(* IEC 61131-3 sources: plcassist-cli/packages/volt-lsp-iec/test-corpus/lenze-mid/Device/Plc Logic/Application/Library Manager/L_CT1P_ControlToolbox, 48 files *)

(* ---- L_CT1P_CONSTANTS.gvl ---- *)
VAR_GLOBAL
	GCWFRICTIONHISTMAX : WORD := 99;
	GCMAXPARITEMS : WORD := 35;
	GCPARITEMSUSED : WORD := 34;
END_VAR

(* ---- L_CT1P_INTERNALCONST.gvl ---- *)
VAR_GLOBAL
END_VAR

(* ---- L_CT1P_IKINAUTOTUNINGEXTERNAL.itf ---- *)
INTERFACE L_CT1P_IKINAUTOTUNINGEXTERNAL
END_INTERFACE

METHOD CALLDEVICEPARAMMANAGERSLAVE
VAR_INPUT
	ECOMMAND : WORD;
	WREGISTERPOSITION : WORD;
	XEXECUTE : BOOL;
END_VAR
VAR_OUTPUT
	XBUSY : BOOL;
	XDONE : BOOL;
	XERROR : BOOL;
	EERRORID : L_Ie1P_Error;
END_VAR
END_METHOD

METHOD CALLMONITORING : BOOL
VAR_INPUT
	XENABLE : BOOL;
END_VAR
END_METHOD

METHOD CHECKPRECONDITIONS : WORD
VAR_INPUT
	XENABLE : BOOL;
	PSCAUTOTUNINGDATAMAININ : POINTER TO BYTE;
END_VAR
END_METHOD

METHOD CLOSEBRAKESPEEDINDEPENDET
VAR_INPUT
	XCLOSBRAKESPEEDINDEPENDET : BOOL;
END_VAR
END_METHOD

METHOD GETMAINFOLLOWERAXIS
VAR_OUTPUT
	PMAINAXISOUT : POINTER TO AXIS_REF;
	PFOLLOWINGAXISOUT : POINTER TO AXIS_REF;
END_VAR
END_METHOD

METHOD SPEEDEQUALSZERO : BOOL
END_METHOD

METHOD STORESAMPLEDBRAKETORQUE
VAR_INPUT
	XSTOREVALUE : BOOL;
END_VAR
END_METHOD

(* ---- _TXERROR.fun ---- *)
FUNCTION _TXERROR : L_IE1P_Error
VAR_INPUT
	WERRCODE : WORD;
END_VAR
END_FUNCTION

(* ---- GETBOOLEANPROPERTY.fun ---- *)
FUNCTION GETBOOLEANPROPERTY : BOOL
VAR_INPUT
	STKEY : WSTRING;
END_VAR
END_FUNCTION

(* ---- GETCOMPANY.fun ---- *)
FUNCTION GETCOMPANY : WSTRING
END_FUNCTION

(* ---- GETNUMBERPROPERTY.fun ---- *)
FUNCTION GETNUMBERPROPERTY : DINT
VAR_INPUT
	STKEY : WSTRING;
END_VAR
END_FUNCTION

(* ---- GETTEXTPROPERTY.fun ---- *)
FUNCTION GETTEXTPROPERTY : WSTRING
VAR_INPUT
	STKEY : WSTRING;
END_VAR
END_FUNCTION

(* ---- GETTEXTPROPERTY2.fun ---- *)
FUNCTION GETTEXTPROPERTY2 : POINTER TO WSTRING
VAR_INPUT
	STKEY : WSTRING;
END_VAR
END_FUNCTION

(* ---- GETTITLE.fun ---- *)
FUNCTION GETTITLE : WSTRING
END_FUNCTION

(* ---- GETVERSION.fun ---- *)
FUNCTION GETVERSION : VERSION
END_FUNCTION

(* ---- GETVERSIONPROPERTY.fun ---- *)
FUNCTION GETVERSIONPROPERTY : VERSION
VAR_INPUT
	STKEY : WSTRING;
END_VAR
END_FUNCTION

(* ---- L_CT1P_CA_CALCDISTANCE.fun ---- *)
FUNCTION L_CT1P_CA_CALCDISTANCE : BOOL
VAR_INPUT
	LRCONSTVELTIME : LREAL;
	LRVELOCITYMAX : LREAL;
	LRACCDECMAX : LREAL;
END_VAR
VAR_OUTPUT
	XERROR : BOOL;
	EERRORID : L_IE1P_Error;
	LRTARGETPOSRELATIVEINT : LREAL;
END_VAR
END_FUNCTION

(* ---- L_CT1P_CA_CALCPROFILEPARAMS.fun ---- *)
FUNCTION L_CT1P_CA_CALCPROFILEPARAMS : BOOL
VAR_INPUT
	LRMAXVELOCITYIN : LREAL := 0;
	LRMAXACCELERATIONIN : LREAL := 0;
	LRMAXDISTANCEIN : LREAL := 0;
END_VAR
VAR_OUTPUT
	LRVELOCITYACTIVE : LREAL := 0;
	LRACCELERATIONACTIVE : LREAL := 0;
	LRMOVEMENTDISTANCEMIN : LREAL := 0;
	LRMOVEMENTDISTANCEMAX : LREAL := 0;
	LRCONSTVELTIME : LREAL := 0;
END_VAR
END_FUNCTION

(* ---- L_CT1P_CA_GETTIMINGOFEXTERNALENCODER.fun ---- *)
FUNCTION L_CT1P_CA_GETTIMINGOFEXTERNALENCODER : BOOL
VAR_OUTPUT
	LRDELAYACTPOS : LREAL;
	LRFILTERCYCLESACTPOS : LREAL;
END_VAR
VAR_IN_OUT
	REALAXIS : _Axis_Ref_Real;
END_VAR
END_FUNCTION

(* ---- L_CT1P_CHECKBASEVALUES.fun ---- *)
FUNCTION L_CT1P_CHECKBASEVALUES : WORD
VAR_INPUT
	PSCCOREDATA : POINTER TO L_CT1P_CA_DeviceParamList;
END_VAR
VAR_IN_OUT
	AXIS : AXIS_REF;
END_VAR
END_FUNCTION

(* ---- L_CT1P_GETOCCOMPDELTAPOSITION.fun ---- *)
FUNCTION L_CT1P_GETOCCOMPDELTAPOSITION : LREAL
VAR_INPUT
	LREIGENFREQ : LREAL;
	LRAMPRATIO : LREAL;
	ECOMPMODE : L_CT1P_OscCompMode;
	LRTARGETVELOCITY : LREAL;
END_VAR
END_FUNCTION

(* ---- L_CT1P_GETOCCOMPDELTATIME.fun ---- *)
FUNCTION L_CT1P_GETOCCOMPDELTATIME : LREAL
VAR_INPUT
	LREIGENFREQ : LREAL;
	ECOMPMODE : L_CT1P_OscCompMode;
END_VAR
END_FUNCTION

(* ---- GLOBALTEXTLIST.fb ---- *)
FUNCTION_BLOCK GLOBALTEXTLIST
VAR
	M_TEXTLISTFILE : STRING(255);
	_STNAMESPACE : STRING;
END_VAR
END_FUNCTION_BLOCK

(* ---- IMAGEPOOL.fb ---- *)
FUNCTION_BLOCK IMAGEPOOL
VAR
	M_STNAMESPACE : STRING(80);
	M_STHELPVARID : STRING;
	M_STHELPVARPATH : STRING(255);
	M_STHELP : STRING;
	M_REGISTERIMAGES : BOOL := TRUE;
END_VAR
END_FUNCTION_BLOCK

METHOD FB_INIT : BOOL
VAR_INPUT
	BINITRETAINS : BOOL;
	BINCOPYCODE : BOOL;
END_VAR
END_METHOD

METHOD FB_REINIT : BOOL
END_METHOD

METHOD FB_EXIT : BOOL
VAR_INPUT
	BINCOPYCODE : BOOL;
END_VAR
END_METHOD

(* ---- L_CT1P_AT_TON.fb ---- *)
FUNCTION_BLOCK L_CT1P_AT_TON
VAR_INPUT
	IN : BOOL;
	PT : TIME;
	LRCYCLE : LREAL;
END_VAR
VAR_OUTPUT
	Q : BOOL;
	ET : TIME;
END_VAR
VAR
	TON_INT : TON;
	TCYLCE : TIME;
	XNOTFIRSTCYCLE : BOOL := FALSE;
END_VAR
END_FUNCTION_BLOCK

(* ---- L_CT1P_AUTOTUNING.fb ---- *)
FUNCTION_BLOCK L_CT1P_AUTOTUNING EXTENDS L_MC1P_Template
VAR_INPUT
	XENABLE : BOOL := FALSE;
	XABORT : BOOL := FALSE;
	XRESETERROR : BOOL := FALSE;
	XEXECUTEIDENT : BOOL := FALSE;
	XENABLEPOSITIONWINDOW : BOOL := FALSE;
	LRPOSITIONWINDOWNEG : LREAL := 1.0;
	LRPOSITIONWINDOWPOS : LREAL := 1.0;
	LRVELOCITYLIMIT : LREAL := 0.0;
	LRACCELERATIONLIMIT : LREAL := 0.0;
	LRDISTANCE : LREAL := 0;
	XRESTOREPARAM : BOOL := FALSE;
	XUSEAXISPARAMETER : BOOL := FALSE;
	EALLOWEDDIRECTION : L_MC1P_ServiceDirection := L_MC1P_ServiceDirection.both;
END_VAR
VAR_OUTPUT
	XERROR : BOOL := FALSE;
	XWARNING : BOOL := FALSE;
	EERRORID : L_IE1P_Error := L_IE1P_Error.NoError;
	XABORTED : BOOL := FALSE;
	XIDENTBUSY : BOOL := FALSE;
	XIDENTDONE : BOOL := FALSE;
	EIDENTIFICATIONSTATE : L_CT1P_CA_IdentificationState := L_CT1P_CA_IdentificationState.PLC_Reset;
	XPOSITIONWINDOWENABLED : BOOL := FALSE;
	LRMVMTVELMAX : LREAL := 0.0;
	LRMVMTACCMAX : LREAL := 0.0;
	LRMVMTDISTANCEMIN : LREAL := 0;
	LRVPNACT : LREAL := 0.0;
	LRTNNACT : LREAL := 0.0;
	LRVPPACT : LREAL := 0.0;
END_VAR
VAR
	RTRESTOREPARAM : R_TRIG;
	EACTSTATE : DWORD := 0;
	XLEAVESERVICESTATE : BOOL := FALSE;
	XDISABLESEEN : BOOL := FALSE;
	XABORTSEEN : BOOL := FALSE;
	XRESETERROROLD : BOOL;
	WCNT : WORD := 0;
	SCCOREDATA : L_CT1P_CA_CoreData := STRUCT(pFB_Par := ADR(fb_InternalParamFB), pFB_AxisReadError := ADR(fb_ReadError), pFB_AxisPower := ADR(fb_Power), pFB_Autotuning := THIS);
	TONAUTOTUNINGDURATION : L_CT1P_AT_TON := STRUCT(PT := TIME#1440m0s0ms);
	XEVENTEXTERNALPARAMFBACTIVATED : BOOL := FALSE;
	LRVELOCITYLIMITINT : LREAL := 0;
	LRACCELERATIONLIMITINT : LREAL := 0;
	LRDISTANCEINT : LREAL := 0;
	XEXECUTEIDENTOLD : BOOL := FALSE;
	DEVICEPARAMMANAGER : L_CT1P_CA_DeviceParamManager;
	PROFILEGENERATOR : L_CT1P_CA_ProfileGenerator;
	MONITORING : L_CT1P_CA_Monitoring;
	QUALITYCRITERIA : L_CT1P_CA_QualityCriteria;
	CHECKPRECONDITIONS : L_CT1P_CA_CheckPreconditions;
	PERFORMAUTOTUNING : L_CT1P_CA_PerformAutotuning;
	FB_READERROR : MC_ReadAxisError;
	FB_POWER : mc_power;
	FB_INTERNALPARAMFB : L_CT1P_ParAutoTuninginternal;
	PAXISREAL : POINTER TO _Axis_Ref_Real;
	PBRAKE : POINTER TO L_MC1P_BrakeControlBase;
	PREALAXIS : POINTER TO _AXIS_REF_COM := 0;
	XWARNINGOLD : BOOL := FALSE;
	LRIMPROVEMENTFACTOR : LREAL := 0;
	XDEACTIVATEERRORINAXIS : BOOL := FALSE;
	EALLOWEDDIRECTIONINT : L_MC1P_ServiceDirection := L_MC1P_ServiceDirection.both;
	TON_MAGNETISATION : L_CT1P_AT_TON;
	XAUTOTUNINGWASACTIVE : BOOL;
	XNEWSTEPENTRY : BOOL;
	ENEWSTATE : DWORD;
	XABORTEDOLD : BOOL;
	ITFKINAUTOTUNING : L_CT1P_IKinAutoTuningExternal;
	STATUSOLD : BOOL;
	XSERVICESTATESETBYAXISCMD : BOOL;
	SERVICESTATESETBYAXISCMND : BOOL;
END_VAR
END_FUNCTION_BLOCK

METHOD ATGETACCELERATION : LREAL
VAR_INPUT
	LRVELOCITY : LREAL := 0;
	LRACCELERATION : LREAL := 0;
END_VAR
VAR_IN_OUT
	AXIS : AXIS_REF;
END_VAR
END_METHOD

METHOD ATGETVELOCITY : LREAL
VAR_INPUT
	LRVELOCITY : LREAL := 0;
	LRVELOTIYRATIOPCT : LREAL := 0;
END_VAR
VAR_IN_OUT
	AXIS : AXIS_REF;
END_VAR
END_METHOD

METHOD CALCULATEIMPROVEMENTFACTOR : LREAL
END_METHOD

METHOD CALLINNERFBINSTANCES
END_METHOD

METHOD CALLMOTIONBLOCKS
END_METHOD

METHOD COPYINPUTS
VAR_IN_OUT
	AXIS : Axis_Ref;
END_VAR
END_METHOD

METHOD SETEXTERNALAUTOTUNINGITF
VAR_INPUT
	PIKINAUTOTUNINGIN : POINTER TO L_CT1P_IKinAutoTuningExternal;
END_VAR
END_METHOD

METHOD STATEMACHINE
END_METHOD

METHOD _GETLIBVERSIONASSTRING : STRING
END_METHOD

METHOD _SETEXTERNALPARAMFB
VAR_INPUT
	PPARAMFB : POINTER TO L_CT1P_ParAutoTuninginternal;
END_VAR
END_METHOD

METHOD STATE_CHECKPRECONDITIONSFOLLOWINGAXIS : DWORD
VAR_INPUT
	XSTOP : BOOL;
	EACTSTATE : DWORD;
	ENEXTSTATE : DWORD;
	EABORTSTATE : DWORD;
	EERRORSTATE : DWORD;
END_VAR
END_METHOD

METHOD STATE_CHECKPRECONDITIONS : DWORD
VAR_INPUT
	XSTOP : BOOL;
	EACTSTATE : DWORD;
	ENEXTSTATE : DWORD;
	EABORTSTATE : DWORD;
	EERRORSTATE : DWORD;
END_VAR
END_METHOD

METHOD STATE_DOAUTOTUNE : DWORD
VAR_INPUT
	XSTOP : BOOL;
	EACTSTATE : DWORD;
	ENEXTSTATE : DWORD;
	EABORTSTATE : DWORD;
	EERRORSTATE : DWORD;
END_VAR
END_METHOD

METHOD STATE_FINISH : DWORD
VAR_INPUT
	XSTOP : BOOL;
	EACTSTATE : DWORD;
	ENEXTSTATE : DWORD;
	EABORTSTATE : DWORD;
	EERRORSTATE : DWORD;
END_VAR
END_METHOD

METHOD STATE_PARAMETERHANDLING : DWORD
VAR_INPUT
	XSTOP : BOOL;
	EACTSTATE : DWORD;
	ENEXTSTATE : DWORD;
	EABORTSTATE : DWORD;
	EERRORSTATE : DWORD;
END_VAR
END_METHOD

(* ---- L_CT1P_AXISCOMMAND_AUTOTUNING.fb ---- *)
FUNCTION_BLOCK L_CT1P_AXISCOMMAND_AUTOTUNING EXTENDS L_MC1P_AxisCommand
VAR_INPUT
	PAXIS : POINTER TO AXIS_REF;
END_VAR
VAR
	FB_AUTOTUNING : L_CT1P_Autotuning;
	SCPARAUTOTUNING : REFERENCE TO L_MC1P_AutotuningPara;
	LRCONSTVELTIME : LREAL := 0;
	LRVELOCITYACTIVE : LREAL := 0;
	LRACCELERATIONACTIVE : LREAL := 0;
	LRDISTANCEACTIVE : LREAL := 0;
	SCPARAUTOTUNING_DUMMY : L_MC1P_AutotuningPara;
	PCONNECTOR : POINTER TO IoConfigConnector;
	ITFAXISCOMMMANDAUTOTUNING : L_MC1P_IAxisCommmand_Autotuning;
	AT_FINISHSTATETEMP : WORD := 0;
	EERRORIDTMP : L_IE1P_error := L_IE1P_Error.NoError;
	WMODULETYPE : UINT;
	XDISABLESET : BOOL := FALSE;
	DWINSTANCE : UDINT;
	WNBOFTUNINGDONE : WORD := 1;
	WNBOFEXPECTEDTUNINGS : WORD := 1;
	LRIMPROVEMENTFACTORSTORED : LREAL;
	PBATEXTERNALITF : POINTER TO BYTE;
	PACTIVEAUTOTUNINGAXIS : ARRAY [1..2] OF POINTER TO _AXIS_REF_REAL;
	C_CMDWORKING10 : USINT := 10;
	C_CMDWORKING30 : USINT := 30;
	C_CMDWORKING50 : USINT := 50;
	C_CMDWORKING70 : USINT := 70;
	C_CMDINVALIDTASKCYCLETIME : USINT := 101;
	C_CMDFUNCTIONNOTSUPPORTEDBYFWVERSION : USINT := 104;
	C_CMDPDOINTERFACEDISABLED : USINT := 106;
	C_CMDTESTMODEALREADYACTIVE : USINT := 107;
	C_CMDINVALIDMOTORCONTROLMODE : USINT := 108;
	C_CMDNOVALIDDIRECTION : USINT := 109;
	C_CMDINSTABILITYWITHCHOSENSTRATEGY : USINT := 110;
	C_CMDAXISNOTHOMED : USINT := 111;
	C_AT_STATE_NOTSTARTED : WORD := 0;
	C_AT_STATE_INITIALIZATION : WORD := 1;
	C_AT_STATE_BACKUPDEVICEPARAM : WORD := 2;
	C_AT_STATE_CHECKPRECONDITIONS : WORD := 3;
	C_AT_STATE_AUTOTUNEVPN : WORD := 4;
	C_AT_STATE_AUTOTUNETNN : WORD := 5;
	C_AT_STATE_AUTOTUNEVPP : WORD := 6;
	C_AT_STATE_FINISHED_1 : WORD := 10;
	C_AT_STATE_FINISHED_2 : WORD := 11;
	C_AT_STATE_FINISHED_3 : WORD := 12;
	C_AT_STATE_BACKUPDEVICEPARAMFOLLOWER : WORD := 22;
	C_AT_STATE_CHECKPRECONDITIONSFOLLOWER : WORD := 23;
	C_AT_STATE_AUTOTUNEVPNFOLLOWER : WORD := 24;
	C_AT_STATE_AUTOTUNETNNFOLLOWER : WORD := 25;
	C_AT_STATE_AUTOTUNEVPPFOLLOWER : WORD := 26;
	C_AT_STATE_FINISHED_4 : WORD := 30;
	C_AT_STATE_FINISHED_5 : WORD := 31;
	C_AT_STATE_FINISHED_6 : WORD := 32;
	C_AT_STATE_FINISHED_7 : WORD := 33;
	C_AT_STATE_FINISHED_8 : WORD := 34;
	C_AT_STATE_FINISHED_9 : WORD := 35;
	C_AT_STATE_ABORTING : WORD := 7;
	C_AT_STATE_ABORTEDBYERROR : WORD := 8;
	C_AT_STATE_ABORTEDBYUSER : WORD := 9;
END_VAR
END_FUNCTION_BLOCK

METHOD ABORTING
END_METHOD

METHOD CALCPROFILEPARAMS
VAR_IN_OUT
	AXIS : AXIS_REF;
END_VAR
END_METHOD

METHOD CALCSTATUS
VAR_IN_OUT
	AXIS : _AXIS_REF_REAL;
END_VAR
END_METHOD

METHOD EXECUTE
END_METHOD

METHOD INITIALIZE : UDINT
VAR_INPUT
	WMODULETYPE : UINT;
	DWINSTANCE : UDINT;
	PCONNECTOR : POINTER TO IoConfigConnector;
END_VAR
END_METHOD

METHOD READINPUTS
END_METHOD

METHOD RESETSTATUSPARAMETER
END_METHOD

METHOD UPDATEAXISPOINTER
VAR_INPUT
	PAXIS : POINTER TO AXIS_REF;
END_VAR
END_METHOD

METHOD UPDATEPARAINTERFACE
VAR_IN_OUT
	SCPAR : L_MC1P_AutotuningPara;
END_VAR
END_METHOD

METHOD FB_INIT : BOOL
VAR_INPUT
	BINITRETAINS : BOOL;
	BINCOPYCODE : BOOL;
END_VAR
END_METHOD

(* ---- L_CT1P_BACKLASHCOMP.fb ---- *)
FUNCTION_BLOCK L_CT1P_BACKLASHCOMP EXTENDS L_MC1P_CompensationBase
VAR_INPUT
	LRBACKLASHWIDTH : LREAL := 0.0;
	LRCOMPTIME : LREAL := 0.1;
	ECOMPMODE : L_CT1P_BacklashCompMode := L_CT1P_BacklashCompMode.NegativeComp;
END_VAR
VAR_OUTPUT
	ECONTACTSTATE : L_CT1P_BacklashContactState := L_CT1P_BacklashContactState.Unknown;
END_VAR
VAR
	FBRAMPGEN : L_MC1P_RampGenerator;
	LRBACKLASHWIDTHINT : LREAL;
	LRCOMPTIMEINT : LREAL;
	ECOMPMODEINT : L_CT1P_BacklashCompMode;
	ECOMPREFERENCEINT : L_CT1P_BacklashCompReference;
	LRACCRATIOINT : LREAL := 0.3333333333;
	ECONTACTSTATEINT : L_CT1P_BacklashContactState;
	LRBACKLASHTARGET : LREAL;
	LRBACKLASHTARGETOLD : LREAL;
	LRBACKLASHPOSACT : LREAL;
	LRBACKLASHVELACT : LREAL;
	LRBACKLASHACCACT : LREAL;
	LRBACKLASHPOSOLD : LREAL;
	LRBACKLASHVELOLD : LREAL;
	LRHOMINGOFFSETACT : LREAL;
	LRENABLEPOS : LREAL;
	LRENABLEDIST : LREAL;
	LRENABLEDISTOLD : LREAL;
	LRVELMAX : LREAL;
	LRACCMAX : LREAL;
	ECOMPREFERENCE : L_CT1P_BacklashCompReference := L_CT1P_BacklashCompReference.SetVelocity;
	_CUSTOMINPUTDATA : ARRAY [1..2] OF L_CT1P_BacklashCompInput;
	_CUSTOMOUTPUTDATA : ARRAY [1..2] OF L_CT1P_BacklashCompOutput;
	_PCUSTOMINPUTDATA : POINTER TO L_CT1P_BacklashCompInput;
	_PCUSTOMOUTPUTDATA : POINTER TO L_CT1P_BacklashCompOutput;
	LRACCRATIO : LREAL;
END_VAR
END_FUNCTION_BLOCK

METHOD CALLCYCLIC2
VAR_IN_OUT
	AXIS : Axis_REf;
END_VAR
END_METHOD

METHOD READINPUTS2
VAR_IN_OUT
	AXIS : Axis_REF;
END_VAR
END_METHOD

METHOD RESETOUTPUTS2
VAR_IN_OUT
	AXIS : Axis_REf;
END_VAR
END_METHOD

METHOD CALCULATE2
VAR_IN_OUT
	AXIS : AXIS_REF;
END_VAR
END_METHOD

METHOD CHECKINPUTDATA2
VAR_IN_OUT
	AXIS : Axis_Ref;
END_VAR
END_METHOD

METHOD ENABLEINIT2
VAR_IN_OUT
	AXIS : Axis_REf;
END_VAR
END_METHOD

METHOD LOADOFFSET2
VAR_INPUT
	OFFSET : LREAL;
END_VAR
VAR_IN_OUT
	AXIS : Axis_REf;
END_VAR
END_METHOD

METHOD GETOFFSETVALUES
VAR_OUTPUT
	LROFFSETPOS : LREAL;
	LROFFSETVEL : LREAL;
	LROFFSETACC : LREAL;
END_VAR
END_METHOD

METHOD CALLFUNCTION
VAR_INPUT
	UIINPUTDATAIDX : UINT;
	UIOUTPUTDATAIDX : UINT;
END_VAR
END_METHOD

METHOD COPYINPUTS : BOOL
VAR_INPUT
	IDX : WORD;
END_VAR
END_METHOD

METHOD COPYOUTPUTS : BOOL
VAR_INPUT
	IDX : WORD;
END_VAR
END_METHOD

METHOD GETCOMPTARGET : LREAL
VAR_INPUT
	LRACTBACKLASHTARGET : LREAL;
END_VAR
VAR_IN_OUT
	AXIS : AXIS_REF;
END_VAR
END_METHOD

METHOD GETCONTACTSTATE : L_CT1P_BacklashContactState
VAR_INPUT
	LRBACKLASHWIDTH : LREAL;
	LRBACKLASHPOSACT : LREAL;
	EACTCONTACTSTATE : L_CT1P_BacklashContactState;
END_VAR
VAR_IN_OUT
	AXIS : AXIS_REF;
END_VAR
END_METHOD

METHOD GETDISTANCESINCEENABLE : LREAL
VAR_IN_OUT
	AXIS : AXIS_REF;
END_VAR
END_METHOD

METHOD GETRAMPPARS : BOOL
VAR_INPUT
	LRCOMPTIME : LREAL;
	LRACCRATIO : LREAL;
	LRBACKLASHWIDTH : LREAL;
END_VAR
VAR_OUTPUT
	LRVELMAX : LREAL;
	LRACCMAX : LREAL;
END_VAR
END_METHOD

METHOD GETTRANSDIR : INT
VAR_IN_OUT
	AXIS : AXIS_REF;
END_VAR
END_METHOD

METHOD INITIALIZEFILTER : BOOL
END_METHOD

(* ---- L_CT1P_CA_CHECKPRECONDITIONS.fb ---- *)
FUNCTION_BLOCK L_CT1P_CA_CHECKPRECONDITIONS
VAR_INPUT
	XEXECUTE : BOOL := FALSE;
	XSTOP : BOOL := FALSE;
	RSCCOREDATA : REFERENCE TO L_CT1P_CA_CoreData;
	RDEVICEPARAMMANAGER : REFERENCE TO L_CT1P_CA_DeviceParamManager;
END_VAR
VAR_OUTPUT
	XBUSY : BOOL := FALSE;
	XDONE : BOOL := FALSE;
	XERROR : BOOL := FALSE;
	EERRORID : L_IE1P_Error := L_IE1P_Error.NoError;
END_VAR
VAR_IN_OUT
	AXIS : AXIS_REF;
END_VAR
VAR
	LRSPEEDFILTERTIME : LREAL;
	LRMOTORINERTIA : LREAL;
	LRLOADINERTIA : LREAL;
	RSCACTPARAM : REFERENCE TO L_CT1P_CA_DeviceParam;
	LRVPPREFERENCEVALUE : LREAL;
	LRDELAYACTPOS : LREAL;
	LRFILTERCYCLESACTPOS : LREAL;
	PREALAXIS : POINTER TO _Axis_Ref_Real;
	REALAXIS : REFERENCE TO _Axis_Ref_Real;
	PBRAKE : POINTER TO L_MC1P_BrakeControlBase;
	XSTOPSEEN : BOOL := FALSE;
	XENABLEPROFILECHECK : BOOL;
	DWSTEP : DWORD := 0;
	RTEXECUTE : R_TRIG;
	PROFILECHECK : L_CT1P_CA_ProfileCheck;
END_VAR
END_FUNCTION_BLOCK

METHOD CALLPROFILECHECK
END_METHOD

METHOD CHECKSTOPELSEPROCEEDWITHSTEP
VAR_INPUT
	DWSTEPINP : DWORD;
END_VAR
END_METHOD

METHOD CHECKVALUES : WORD
VAR_IN_OUT
	AXIS : AXIS_REF;
END_VAR
END_METHOD

METHOD RAISEERROR
VAR_INPUT
	ERRCODE : L_IE1P_Error;
END_VAR
END_METHOD

METHOD RAISEFINISHED
END_METHOD

METHOD RAISESTOP
END_METHOD

METHOD READWRITEVALUES : WORD
VAR_IN_OUT
	DWSTEP : DWORD;
	AXIS : AXIS_REF;
END_VAR
END_METHOD

METHOD RESET : BOOL
END_METHOD

METHOD STATEMACHINE
END_METHOD

(* ---- L_CT1P_CA_DEVICEPARAMMANAGER.fb ---- *)
FUNCTION_BLOCK L_CT1P_CA_DEVICEPARAMMANAGER
VAR_INPUT
	ECOMMAND : L_CT1P_CA_DPMCommand := L_CT1P_CA_DPMCommand.None;
	RSCPARAMLIST : REFERENCE TO L_CT1P_CA_DeviceParamList;
	WREGISTERPOSITION : WORD;
	XEXECUTE : BOOL := FALSE;
END_VAR
VAR_OUTPUT
	XBUSY : BOOL := FALSE;
	XDONE : BOOL := FALSE;
	XERROR : BOOL := FALSE;
	EERRORID : L_Ie1P_Error;
END_VAR
VAR_IN_OUT
	AXIS : Axis_ref;
END_VAR
VAR
	WRITEPARAMETER : MC_WriteParameter;
	READPARAMETER : MC_ReadParameter;
	PDCOREAD : POINTER TO L_MC1P.L_DCO_ReadDriveParameter;
	PDCOWRITE : POINTER TO L_MC1P.L_DCO_WriteDriveParameter;
	WWRITEMODE : WORD;
	ECOMMANDINT : L_CT1P_CA_DPMCommand := L_CT1P_CA_DPMCommand.None;
	WREGISTERPOSITIONINT : WORD;
	WIDX : WORD := 1;
	WIDX2 : WORD := 1;
	XEXECUTEOLD : BOOL;
	XINITIALVALUESREADED : BOOL;
	XSUSPENDERRORMESSAGE : BOOL;
	APARAMCHANGED : ARRAY [1..L_Ct1P_Constants.gcMaxParItems] OF BOOL;
	PREALAXIS : POINTER TO _AXIS_REF_REAL;
	XBUSYKIN : BOOL;
	XDONEKIN : BOOL;
	XERRORKIN : BOOL;
	EERRORIDKIN : L_IE1P_Error;
	XBUSYINT : BOOL;
	XDONEINT : BOOL;
	XERRORINT : BOOL;
	EERRORIDINT : L_IE1P_Error;
	PATDATAFOLLOWINGAXIS : POINTER TO L_CT1P_CA_DeviceParamList;
	ITFKINAUTOTUNING : L_CT1P_IKinAutoTuningExternal;
	KINAUTOTUNING : L_CT1P_IKinAutoTuningExternal;
END_VAR
END_FUNCTION_BLOCK

METHOD CHECKERRORS
VAR_IN_OUT
	AXIS : Axis_Ref;
END_VAR
END_METHOD

METHOD READ : BOOL
VAR_INPUT
	RSCPARAM : REFERENCE TO L_CT1P_CA_DeviceParam;
END_VAR
VAR_IN_OUT
	AXIS : Axis_Ref;
END_VAR
END_METHOD

METHOD RESETOUTPUTS
END_METHOD

METHOD STOREINPUTS
END_METHOD

METHOD STOREPARAMSPERSISTENT : BOOL
VAR_IN_OUT
	AXIS : Axis_Ref;
END_VAR
END_METHOD

METHOD WRITE : BOOL
VAR_INPUT
	RSCPARAM : REFERENCE TO L_CT1P_CA_DeviceParam;
END_VAR
VAR_IN_OUT
	AXIS : Axis_Ref;
END_VAR
END_METHOD

(* ---- L_CT1P_CA_MONITORING.fb ---- *)
FUNCTION_BLOCK L_CT1P_CA_MONITORING
VAR_INPUT
	XENABLE : BOOL := FALSE;
	RSCCOREDATA : REFERENCE TO L_CT1P_CA_CoreData;
END_VAR
VAR_OUTPUT
	XAXISDISABLED : BOOL := FALSE;
	XAXISERROR : BOOL := FALSE;
	XPOSLIMITMINEXCEEDED : BOOL := FALSE;
	XPOSLIMITMAXEXCEEDED : BOOL := FALSE;
	XINSTABILITYBYCONTROLLERCONSTRAINTS : BOOL := FALSE;
	XINSTABILITYBYFREQUENCYANALYSIS : BOOL := FALSE;
	XINSTABILITYBYVELOCITYOVERSHOOT : BOOL := FALSE;
END_VAR
VAR_IN_OUT
	AXIS : AXIS_REF;
END_VAR
VAR
	TONAXISISDISABLED : L_CT1P_AT_TON;
	AXINSTABILITYBUFFER : ARRAY [0..9] OF BOOL;
	XVALID : BOOL := FALSE;
	XINIT : BOOL := FALSE;
	TEOFWTMP : BOOL := FALSE;
	XPOSCTRLLIMITED : BOOL;
	XINSTABILITYEXTERNAL : BOOL;
	BBUFFER : BYTE;
	WINSTABILITYBUFFERINDEX : WORD := 0;
	WINDEX : WORD := 0;
	WTRUECOUNT : WORD := 0;
	WBUFFER1 : WORD;
	WCNT : WORD := 0;
	WXNCNT2 : WORD := 0;
	DIPARAM : DINT;
	LRVELERROR : LREAL := 0;
	PREALAXIS : POINTER TO _Axis_Ref_Real;
	REALAXIS : REFERENCE TO _Axis_Ref_Real;
	MC_READINSTABILITY : MC_ReadParameter;
	PDCOREAD : POINTER TO L_MC1P.L_DCO_ReadDriveParameter;
	LRPSI2 : LREAL := 0;
	ALRXN2 : ARRAY [0..7] OF LREAL;
	LRFILTERINPUT1MS : LREAL;
	LRFILTERINPUT10MS : LREAL;
	PT1256MS : L_USPP_PT1Filter;
	PT1256MS_10 : L_USPP_PT1Filter;
	STEOVALUES10MS : L_CT1P_TEOValues;
	STEOVALUES1MS : L_CT1P_TEOValues;
	ALRELLIPVALUESIN : ARRAY [0..7] OF LREAL;
	ALRELLIPTVALUESOUT : ARRAY [0..7] OF LREAL;
	ITFKINAUTOTUNING : L_CT1P_IKinAutoTuningExternal;
	CWTEODEPTHMAX : WORD := 7;
	KINAUTOTUNING : L_CT1P_IKinAutoTuningExternal;
	STIMULATEINSTABILITY : BOOL;
END_VAR
END_FUNCTION_BLOCK

METHOD ELLIPTICFILTER : LREAL
VAR_INPUT
	LRIN : LREAL;
	XRESET : BOOL;
END_VAR
VAR_IN_OUT
	ALRELLIPVALUESIN : ARRAY [0..7] OF LREAL;
	ALRELLIPVALUESOUT : ARRAY [0..7] OF LREAL;
	BBUFFER : BYTE;
END_VAR
END_METHOD

METHOD MAIN
VAR_INPUT
	XENABLE : BOOL := FALSE;
	LRTEOLIMIT1 : LREAL;
	LRTEOLIMIT2 : LREAL;
	XISCIAADVANCEDAXIS : BOOL;
	XEXTERNALPOSITIONFEEDBACK : BOOL;
	XAXISENABLEDREAL : BOOL;
	XTEOLIMITVALID : BOOL;
END_VAR
VAR_OUTPUT
	XAXISDISABLED : BOOL := FALSE;
	XAXISERROR : BOOL := FALSE;
	XPOSLIMITMINEXCEEDED : BOOL := FALSE;
	XPOSLIMITMAXEXCEEDED : BOOL := FALSE;
	XINSTABILITYBYCONTROLLERCONSTRAINTS : BOOL := FALSE;
	XINSTABILITYBYFREQUENCYANALYSIS : BOOL := FALSE;
	XINSTABILITYBYVELOCITYOVERSHOOT : BOOL := FALSE;
	XINSTABILITYKIN : BOOL := FALSE;
END_VAR
VAR_IN_OUT
	AXIS : AXIS_REF;
END_VAR
END_METHOD

METHOD TEOFW : BOOL
VAR_IN_OUT
	AXIS : AXIS_REF;
	DIPARAM : DINT;
END_VAR
END_METHOD

METHOD TEOPLCPOSITION : BOOL
VAR_INPUT
	XOPTIMISINGEXTERNALFEEDBACK : BOOL;
	LRVPPACTUALVALUE : LREAL;
END_VAR
VAR_IN_OUT
	AXIS : AXIS_REF;
END_VAR
END_METHOD

METHOD TEAGERENERGYOPERATOR
VAR_INPUT
	LRINPUT : LREAL;
	XRESET : BOOL;
	WCALCULATIONTIME : WORD;
END_VAR
VAR_IN_OUT
	STEOVALUES : L_CT1P_TEOValues;
END_VAR
END_METHOD

(* ---- L_CT1P_CA_PERFORMAUTOTUNING.fb ---- *)
FUNCTION_BLOCK L_CT1P_CA_PERFORMAUTOTUNING
VAR_INPUT
	XEXECAUTOTUNEVPN : BOOL := FALSE;
	XEXECAUTOTUNETNN : BOOL := FALSE;
	XEXECAUTOTUNEVPP : BOOL := FALSE;
	XEXECSTARTMOVEMENT : BOOL := FALSE;
	XSTOP : BOOL := FALSE;
	RSCCOREDATA : REFERENCE TO L_CT1P_CA_CoreData;
	RDEVICEPARAMMANAGER : REFERENCE TO L_CT1P_CA_DeviceParamManager;
	RPROFILEGENERATOR : REFERENCE TO L_CT1P_CA_ProfileGenerator;
	RMONITORING : REFERENCE TO L_CT1P_CA_Monitoring;
	RQUALITYCRITERIA : REFERENCE TO L_CT1P_CA_QualityCriteria;
END_VAR
VAR_OUTPUT
	XBUSY : BOOL := FALSE;
	XDONE : BOOL := FALSE;
	XERROR : BOOL := FALSE;
	EERRORID : L_IE1P_Error := L_IE1P_Error.NoError;
END_VAR
VAR_IN_OUT
	AXIS : AXIS_REF;
END_VAR
VAR
	DWSTEPCOMPLETE : DWORD := 0;
	DWSTEPMAJOR : DWORD := 0;
	DWSTEPMINOR : DWORD := 0;
	RTEXECAUTOTUNEVPN : R_TRIG;
	RTEXECAUTOTUNETNN : R_TRIG;
	RTEXECAUTOTUNEVPP : R_TRIG;
	RTEXECSTARTMOVEMENT : R_TRIG;
	LRQUYLITYCRITERIAMIN : LREAL := 0;
	XPHASE1COMPLETED : BOOL := FALSE;
	XPHASE2COMPLETED : BOOL := FALSE;
	XSTOPSEEN : BOOL := FALSE;
	XPROCEEDWITHPHASE2B : BOOL := FALSE;
	DNPROFILETASKCYCLECOUNT : DINT := 0;
	PAXISREAL : POINTER TO _Axis_Ref_Real;
	PBRAKE : POINTER TO L_MC1P_BrakeControlBase;
	LRINSTABILITYFACTOR : LREAL := 0.45;
	LRSTEPFACTOR_PCT : LREAL := 100;
	XINSTABILITYDETECTED : BOOL := FALSE;
	XIGNOREQUALITY : BOOL := FALSE;
	XOPTIMIZETNN : BOOL := FALSE;
	XAXISPOWERSTATUSOLD : BOOL;
	XMAXPARAMVALUESETTED : BOOL := FALSE;
	XMINPARAMVALUESETTED : BOOL := FALSE;
	XWAITTIMERON : BOOL;
	XWAITTIMERONOLD : BOOL;
	XWAITTIMEREACHED : BOOL;
	XQUALITYCRITERIAENABLEOLD : BOOL;
	XCALCULATELIMITSFORTESTMOTION : BOOL;
	WWAITAFTERINSTABILITY : WORD;
	WIDENTSTEPTMP : WORD;
	WINSTABILITYSTEPS : WORD;
	DWNEXTSTEP : DWORD;
	DWWAITTIMECNTR : WORD;
	WMAXVALUECOUNTER : WORD;
	WMINVALUECOUNTER : WORD;
	WWAITAFTERINSTABILITYINACTIVE : WORD;
	WINSTABLITCNT : WORD;
	DWFIRSTACTIVATIONSTEP : DWORD;
	LRWAITINGTIME : LREAL;
	ALRTNNTEOVALUES : ARRAY [0..2, 0..10] OF LREAL;
	LRTEO1TMP : LREAL;
	LRTEO2TMP : LREAL;
	RSCACTPARAM : REFERENCE TO L_CT1P_CA_DeviceParam;
	LRACTVELOCITYMAXWHILEENABLED : LREAL;
	LRACTTORQUEMAXWHILEENABLED : LREAL;
	TONAXISPOWER : L_CT1P_AT_TON;
	ITFKINAUTOTUNING : L_CT1P_IKinAutoTuningExternal;
	KINAUTOTUNING : L_CT1P_IKinAutoTuningExternal;
END_VAR
END_FUNCTION_BLOCK

METHOD CHECKERRORS : BOOL
VAR_IN_OUT
	AXIS : Axis_Ref;
END_VAR
END_METHOD

METHOD CHECKSTOPELSEPROCEEDWITHFIRSTACTIVATIONSTEP
VAR_INPUT
	DWSTEPINP : DWORD;
END_VAR
END_METHOD

METHOD CHECKSTOPELSEPROCEEDWITHMINORSTEP
VAR_INPUT
	DWSTEPINP : DWORD;
END_VAR
END_METHOD

METHOD HANDLINGTEOLIMITS
END_METHOD

METHOD INITPROFILER
VAR_INPUT
	XMOVETOSTARTPOSITION : BOOL := FALSE;
END_VAR
VAR_IN_OUT
	AXIS : AXIS_REF;
END_VAR
END_METHOD

METHOD INSTABIITYDETECTED : BOOL
VAR_INPUT
	DWNEXTSTEPIN : DWORD;
	LRINSTABILITYFACTOR : LREAL;
END_VAR
VAR_OUTPUT
	XINSTABILITYDETECTED : BOOL;
END_VAR
VAR_IN_OUT
	AXIS : AXIS_REF;
	RSCACTPARAM : L_CT1P_CA_DeviceParam;
	LRACTUALPARAMVALUE : LREAL;
	LRACTUALSTEPVALUE : LREAL;
	DWNEXTSTEPOUT : DWORD;
	WINSTABILITYSTEPS : WORD;
END_VAR
END_METHOD

METHOD RAISEERROR
VAR_INPUT
	ERRCODE : L_IE1P_Error;
END_VAR
END_METHOD

METHOD RAISEFINISHED
END_METHOD

METHOD RAISESTOP
END_METHOD

METHOD RESET : BOOL
END_METHOD

METHOD STATEMACHINE_FIRSTACTIVATION : BOOL
VAR_IN_OUT
	AXIS : AXIS_REF;
END_VAR
END_METHOD

METHOD STATEMACHINE
END_METHOD

METHOD STATEMACHINE_MAJOR00
END_METHOD

METHOD STATEMACHINE_OPTIMIZING
VAR_IN_OUT
	AXIS : AXIS_REF;
	RSCACTPARAM : L_CT1P_CA_DeviceParam;
	LRACTUALVALUE : LREAL;
	LRSTEPVALUE : LREAL;
END_VAR
END_METHOD

METHOD WAITTIMER : BOOL
VAR_IN_OUT
	AXIS : AXIS_REF;
END_VAR
END_METHOD

METHOD RESETTEOLIMITS
END_METHOD

METHOD SELECTVALUESFORPARAMETER
VAR_IN_OUT
	AXIS : AXIS_REF;
	RSCACTPARAM : L_CT1P_CA_DeviceParam;
END_VAR
END_METHOD

METHOD SETPARAMVALUE
VAR_INPUT
	LRSETVALUE : LREAL;
END_VAR
VAR_IN_OUT
	RSCACTPARAM : L_CT1P_CA_DeviceParam;
END_VAR
END_METHOD

(* ---- L_CT1P_CA_PROFILECHECK.fb ---- *)
FUNCTION_BLOCK L_CT1P_CA_PROFILECHECK
VAR_INPUT
	XENABLE : BOOL := FALSE;
	RSCCOREDATA : REFERENCE TO L_CT1P_CA_CoreData := 0;
	XENABLEPOSITIONWINDOW : BOOL := FALSE;
	LRPOSITIONWINDOWNEG : LREAL := 0.0;
	LRPOSITIONWINDOWPOS : LREAL := 0.0;
	LRVELOCITYLIMIT : LREAL := 0.0;
	LRACCELERATIONLIMIT : LREAL := 0.0;
	LRDISTANCE : LREAL := 0.0;
END_VAR
VAR_OUTPUT
	XBUSY : BOOL := FALSE;
	XDONE : BOOL := FALSE;
	XWARNING : BOOL := FALSE;
	XERROR : BOOL := FALSE;
	EERRORID : L_IE1P_Error := L_IE1P_Error.NoError;
END_VAR
VAR_IN_OUT
	AXIS : AXIS_REF;
END_VAR
VAR
	DWSTEP : DWORD := 0;
	XCHECKNEEDED : BOOL := FALSE;
	XWARNING_LOCAL : BOOL := FALSE;
	XERROR_LOCAL : BOOL := FALSE;
	EERRORID_LOCAL : L_IE1P_Error := L_IE1P_Error.NoError;
	LRSWLIMITMIN : LREAL;
	LRSWLIMITMAX : LREAL;
	PREALAXIS : POINTER TO _AXIS_REF_REAL;
	ETRAVERSINGRANGE_ACT : L_MC1P_TraversingRange := L_MC1P_TraversingRange.Limited;
	XHOMEPOSAVAILABLE_ACT : BOOL := FALSE;
	XSWLIMITENABLED_ACT : BOOL := FALSE;
	XENABLEPOSITIONWINDOW_ACT : BOOL := FALSE;
	LRPOSITIONWINDOWNEG_ACT : LREAL := 0.0;
	LRPOSITIONWINDOWPOS_ACT : LREAL := 0.0;
	LRVELOCITYLIMIT_ACT : LREAL := 0.0;
	LRACCELERATIONLIMIT_ACT : LREAL := 0.0;
	LRDISTANCEMAX_ACT : LREAL := 0.0;
	LRMAXVELOCITYAPPL_ACT : LREAL := 0.0;
	LRMAXACCELERATIONAPPL_ACT : LREAL := 0.0;
	LRSWLIMITNEG_ACT : LREAL := 0.0;
	LRSWLIMITPOS_ACT : LREAL := 0.0;
	LRSCALEUNITTORPM_ACT : LREAL := 0.0;
END_VAR
END_FUNCTION_BLOCK

METHOD RAISEERROR
VAR_INPUT
	ERRCODE : L_IE1P_Error;
END_VAR
END_METHOD

METHOD RAISEFINISHED
END_METHOD

METHOD RAISEWARNING
VAR_INPUT
	ERRCODE : L_IE1P_Error;
END_VAR
END_METHOD

METHOD STATEMACHINE
END_METHOD

(* ---- L_CT1P_CA_PROFILEGENERATOR.fb ---- *)
FUNCTION_BLOCK L_CT1P_CA_PROFILEGENERATOR EXTENDS L_MC1P_Template_IntFB
VAR_INPUT
	XEXECUTE : BOOL;
	XSTOP : BOOL;
	XUSEEXTERNALPOSITION : BOOL := FALSE;
	LRSETPOSRELATIVE : LREAL := 0;
	LRVCONSTDURATION_S : LREAL := 0;
	LRVELOCITYMAX : LREAL;
	LRACCDECMAX : LREAL;
	LRINPOSTIMEOUT : LREAL := 1.0;
	XPOSITIVE : BOOL := TRUE;
	WCYCLECOUNT : WORD;
	LRSTANDSTILLDURATION_S : LREAL;
	XONEDIRECTION : BOOL;
	XREVERSING : BOOL;
	WFUNID : WORD;
END_VAR
VAR_OUTPUT
	XDONE : BOOL;
	XBUSY : BOOL;
	XCOMMANDABORTED : BOOL;
	XERROR : BOOL;
	EERRORID : L_IE1P_Error;
END_VAR
VAR_IN_OUT
	AXIS : Axis_Ref;
END_VAR
VAR
	XFIRSTCYCLE : BOOL;
	XEXECUTEOLD : BOOL;
	XRESETOUTPUT : BOOL;
	XINTERNALABORT : BOOL;
	XUSEEXTERNALPOSITIONINT : BOOL := FALSE;
	XPOSITIVEINT : BOOL;
	WCYCLECOUNTINT : WORD;
	LRSETPOSRELATIVEINT : LREAL;
	LRVELOCITYMAXINT : LREAL;
	LRACCDECMAXINT : LREAL;
	LRINPOSTOLERANCEINT : LREAL := 100.0;
	LRINPOSMAXVELOCITYINT : LREAL := 100;
	LRINPOSTIMEOUTINT : LREAL := 1.0;
	LRSTANDSTILLDURATION_SINT : LREAL;
	LRRELATIVETARGETPOS : LREAL;
	L_MC1P_POSPROFILER1 : REFERENCE TO L_Mc1P_PosProfiler;
	SCPROFILEPARAMETER : L_MC1P_ProfileParameter;
	WPROFILESTATE : WORD;
	WCYCLECOUNTER : WORD;
	DWVALIDCOUNTER : DWORD;
	XSTOPOLD : BOOL;
	XPOSPROFILERINUSE : BOOL;
	XDIRECTIONCHANGE : BOOL;
	XREVERSINGINT : BOOL;
	FBBASE : L_MC1P_Template;
	LRSETPOSINIT : LREAL;
	PREALAXIS : POINTER TO _AXIS_REF_Real;
	LRACTVELOCITYOLD : LREAL;
	LRSTANDSTILLDURATION_ACTIVE : LREAL;
	ITFKINAUTOTUNING : L_CT1P_IKinAutoTuningExternal;
	XKINEQUALYZERO : BOOL;
	FUNCTIONTYPE : L_MC1P_TypeFunction;
	KINAUTOTUNING : L_CT1P_IKinAutoTuningExternal;
	POSPROFILERINUSE : BOOL;
END_VAR
END_FUNCTION_BLOCK

METHOD CHECKPRECONDITION : BOOL
VAR_OUTPUT
	EERRORID : L_IE1P_Error;
END_VAR
END_METHOD

METHOD CYCLIC
VAR_IN_OUT
	AXIS : AXIS_REF;
	FBBASE : L_MC1P_Template;
END_VAR
END_METHOD

METHOD INIT
VAR_IN_OUT
	AXIS : AXIS_REF;
	FBBASE : L_MC1P_Template;
END_VAR
END_METHOD

METHOD MAIN
VAR_IN_OUT
	AXIS : AXIS_REF;
	FBBASE : L_MC1P_Template;
END_VAR
END_METHOD

METHOD MOVEMENTPROFILE
VAR_IN_OUT
	AXIS : Axis_ref;
END_VAR
END_METHOD

METHOD RESETOUTPUTS
END_METHOD

METHOD STOREINPUTS
VAR_IN_OUT
	AXIS : AXIS_REF;
END_VAR
END_METHOD

METHOD ABORTACTIVEFUNCTION : BOOL
END_METHOD

METHOD SETINTERNALSTOP : BOOL
VAR_INPUT
	XSTOP : BOOL;
	ESETSTATE : L_MC1P_AXIS_STATE;
	XPOSMODE : BOOL := FALSE;
	LRTARGETPOS : LREAL := 0;
	XABORTACTIVEFUNCTION : BOOL := TRUE;
END_VAR
VAR_IN_OUT
	XSTOPACTIVE : BOOL;
	XSTOPDONE : BOOL;
END_VAR
END_METHOD

(* ---- L_CT1P_CA_QUALITYCRITERIA.fb ---- *)
FUNCTION_BLOCK L_CT1P_CA_QUALITYCRITERIA
VAR_INPUT
	XENABLE : BOOL := FALSE;
	WVALUESELECTION : WORD := 0;
	LRNOMVELOCITY : LREAL := 1.0;
END_VAR
VAR_OUTPUT
	LRSELECTEDVALUESUM : LREAL := 0.0;
	LRVELERRORSUM : LREAL := 0.0;
	LRPOSERRORSUM : LREAL := 0.0;
	LRVELOVERSHOOT_PCT : LREAL := -100.0;
END_VAR
VAR_IN_OUT
	AXIS : AXIS_REF;
END_VAR
VAR
	LRVELOVERSHOOTAVFACTOR : LREAL := 0.8;
	RTENABLE : R_TRIG;
	LRSETVELLASTCYCLE : LREAL := 0.0;
	LRSETPOSLASTCYCLE : LREAL := 0.0;
	LRVELOVERSHOOTACT : LREAL;
	LRVELOVERSHOOTNEW : LREAL;
	WTASKCYCLE_MS : WORD := 1;
	ALRVELERR : ARRAY [0..3] OF LREAL := [0.0, 0.0, 0.0, 0.0];
	PREALAXIS : POINTER TO _AXIS_REF_REAL;
	REALAXIS : REFERENCE TO _AXIS_REF_REAL;
	DWSETVELOCITYSTORESIZE : DWORD := 16;
	ALRSETVELOCITYSTORE : ARRAY [0..dwSetVelocityStoreSize] OF LREAL;
	DWSETVELOCITYWRITEIDX : DWORD := 0;
	DWSETVELOCITYSHIFTFACTOR : DWORD := 3;
	LRSETVELOCITYSHIFTED : LREAL := 0.0;
	LRVELERRORSUMTMP : LREAL := 0;
	LRPOSERRORSUMTMP : LREAL := 0;
	LRVALUECNT : LREAL := 0;
	DWCNT : DWORD := 0;
	PT1_FILTER_ACTVEL : L_USPP_PT1Filter;
END_VAR
END_FUNCTION_BLOCK

(* ---- L_CT1P_CROSSCOMP.fb ---- *)
FUNCTION_BLOCK L_CT1P_CROSSCOMP EXTENDS L_MC1P_CompensationBase
VAR_INPUT
	ALRBASEPOSITION : POINTER TO LREAL;
	ALRAXISCORRECTION : POINTER TO LREAL;
END_VAR
VAR_OUTPUT
	LRACTCORRECTION : LREAL;
END_VAR
VAR_IN_OUT
	BASE : AXIS_REF;
END_VAR
VAR
	LICHANDLING : L_IMHP_LLMHandling;
	FBLININTERP : L_UMTP_InterpolationLinear;
	SCINTERPDATAINT : L_UMTP_InterpolationData;
	LRCORRECTIONPOS : LREAL;
	LRCORRECTIONPOSOLD : LREAL;
	LRCORRECTIONVEL : LREAL;
	LRCORRECTIONVELOLD : LREAL;
	LRCORRECTIONACC : LREAL;
	DINBROFVALUES : DINT;
	XFIRSTCALL : BOOL;
	_CUSTOMINPUTDATA : ARRAY [1..2] OF L_CT1P_CrossCompInput;
	_CUSTOMOUTPUTDATA : ARRAY [1..2] OF L_CT1P_CrossCompOutput;
	_PCUSTOMINPUTDATA : POINTER TO L_CT1P_CrossCompInput;
	_PCUSTOMOUTPUTDATA : POINTER TO L_CT1P_CrossCompOutput;
END_VAR
END_FUNCTION_BLOCK

METHOD CALLCYCLIC2
VAR_IN_OUT
	AXIS : L_MC1P.Axis_REf;
END_VAR
END_METHOD

METHOD CHECKINPUTDATA2
VAR_IN_OUT
	AXIS : Axis_REf;
END_VAR
END_METHOD

METHOD READINPUTS2
VAR_IN_OUT
	AXIS : Axis_REf;
END_VAR
END_METHOD

METHOD RESETOUTPUTS2
VAR_IN_OUT
	AXIS : Axis_REf;
END_VAR
END_METHOD

METHOD CALCULATE2
VAR_IN_OUT
	AXIS : Axis_REf;
END_VAR
END_METHOD

METHOD FILTERSTARTCONDITION
VAR_INPUT
	LRSETPOS : LREAL;
	LRSETVEL : LREAL;
	LRSETACC : LREAL;
END_VAR
VAR_IN_OUT
	AXIS : L_MC1P.Axis_ref;
END_VAR
END_METHOD

METHOD GETOFFSETVALUES
VAR_OUTPUT
	LROFFSETPOS : LREAL;
	LROFFSETVEL : LREAL;
	LROFFSETACC : LREAL;
END_VAR
END_METHOD

METHOD CALLFUNCTION
VAR_INPUT
	UIINPUTDATAIDX : UINT;
	UIOUTPUTDATAIDX : UINT;
END_VAR
END_METHOD

METHOD COPYINPUTS : BOOL
VAR_INPUT
	IDX : WORD;
END_VAR
END_METHOD

METHOD COPYOUTPUTS : BOOL
VAR_INPUT
	IDX : WORD;
END_VAR
END_METHOD

(* ---- L_CT1P_KALMANFILTER_INTERNAL.fb ---- *)
FUNCTION_BLOCK L_CT1P_KALMANFILTER_INTERNAL
VAR_INPUT
	LRT_CYCLEINTERVAL : LREAL;
	LRT_CYCLEINTERVALINV : LREAL;
	LRNORMGK : LREAL := ((100.0 * 60.0) / ((3000.0 * 2) * 3.14159265));
	ALRX0_VALUE : ARRAY [0..4] OF LREAL;
	ALRP : ARRAY [0..24] OF LREAL;
	ALRA : ARRAY [0..24] OF LREAL;
	I : ARRAY [0..24] OF SINT;
	ALRK : ARRAY [0..4] OF LREAL;
	A : ARRAY [0..4] OF LREAL;
	LRJ : LREAL;
	B : LREAL;
	K : DINT;
	ALRA_0 : ARRAY [0..24] OF LREAL;
	B_I : DINT;
	I_0 : DINT;
	RTB_ALRY_IDX : LREAL;
	RTB_ALRY_IDX_1 : LREAL;
	RTB_ALRX : ARRAY [0..4] OF LREAL;
	LRCNT : LREAL;
	LRMW : LREAL;
	ALRXV : ARRAY [0..4] OF LREAL;
	ALRPV : ARRAY [0..24] OF LREAL;
	ALRFELD : ARRAY [0..69] OF LREAL;
	ALRQ_VALUE : ARRAY [0..24] OF LREAL := [1E-05, 0.0, 0.0, 0.0, 0.0, 0.0, 1E-06, 0.0, 0.0, 0.0, 0.0, 0.0, 0.0001, 0.0, 0.0, 0.0, 0.0, 0.0, 0.0001, 0.0, 0.0, 0.0, 0.0, 0.0, 0.0001];
	LRR_VALUE : LREAL := 0.1;
	ALRP_VALUE : ARRAY [0..24] OF LREAL := [1E-05, 0.0, 0.0, 0.0, 0.0, 0.0, 100.0, 0.0, 0.0, 0.0, 0.0, 0.0, 10.0, 0.0, 0.0, 0.0, 0.0, 0.0, 10, 0.0, 0.0, 0.0, 0.0, 0.0, 10];
	LRSCALECOULOMB : LREAL := 100;
	F : ARRAY [0..4] OF SINT := [0, 1, 0, 0, 0];
	E : ARRAY [0..4] OF SINT := [0, 0, 1, 0, 0];
	B_D : ARRAY [0..4] OF SINT := [0, 0, 0, 1, 0];
	C : ARRAY [0..4] OF SINT := [0, 0, 0, 0, 1];
	D_B : ARRAY [0..4] OF SINT := [1, 0, 0, 0, 0];
END_VAR
VAR_OUTPUT
	LRVELOCITYIDENT : LREAL;
	LRINERTIAIDENTKGM2 : LREAL;
	LRVISCOUSDAMPINGIDENT : LREAL;
	LRCONSTANTTORQUEIDENT : LREAL;
	LRIDENTCOULOMBFRICTION : LREAL;
END_VAR
VAR
	LRTORQUEINT : LREAL;
	LRACCINT : LREAL;
END_VAR
END_FUNCTION_BLOCK

METHOD KALMANFILTER : BOOL
VAR_INPUT
	LRM_IST : LREAL;
	LROMEGA_IST : LREAL;
END_VAR
END_METHOD

METHOD KALMANFILTERINITVALUES
END_METHOD

METHOD SETMATRIXVALUESTOIDENTALL : BOOL
END_METHOD

METHOD SETMATRIXVALUESTOIDENTDAMPING : BOOL
END_METHOD

METHOD SETMATRIXVALUESTOIDENTINERTIA : BOOL
END_METHOD

METHOD SETMATRIXVALUESTOIDENTTORQUE : BOOL
END_METHOD

(* ---- L_CT1P_LEADSCREWERRORCOMP.fb ---- *)
FUNCTION_BLOCK L_CT1P_LEADSCREWERRORCOMP EXTENDS L_MC1P_CompensationBase
VAR_INPUT
	ALRAXISPOSITION : POINTER TO LREAL;
	ALRAXISCORRECTION : POINTER TO LREAL;
END_VAR
VAR_OUTPUT
	LRACTCORRECTION : LREAL;
END_VAR
VAR
	LICHANDLING : L_IMHP_LLMHandling;
	FBLININTERP : L_UMTP_InterpolationLinear;
	SCINTERPDATAINT : L_UMTP_InterpolationData;
	LRCORRECTIONPOS : LREAL;
	LRCORRECTIONPOSOLD : LREAL;
	LRCORRECTIONVEL : LREAL;
	LRCORRECTIONVELOLD : LREAL;
	LRCORRECTIONACC : LREAL;
	DINBROFVALUES : DINT;
	XFIRSTCALL : BOOL;
	_CUSTOMINPUTDATA : ARRAY [1..2] OF L_CT1P_LeadscrewErrorCompInput;
	_CUSTOMOUTPUTDATA : ARRAY [1..2] OF L_CT1P_LeadscrewErrorCompOutput;
	_PCUSTOMINPUTDATA : POINTER TO L_CT1P_LeadscrewErrorCompInput;
	_PCUSTOMOUTPUTDATA : POINTER TO L_CT1P_LeadscrewErrorCompOutput;
END_VAR
END_FUNCTION_BLOCK

METHOD CALLCYCLIC2
VAR_IN_OUT
	AXIS : Axis_REf;
END_VAR
END_METHOD

METHOD READINPUTS2
VAR_IN_OUT
	AXIS : Axis_REf;
END_VAR
END_METHOD

METHOD RESETOUTPUTS2
VAR_IN_OUT
	AXIS : Axis_REf;
END_VAR
END_METHOD

METHOD CALCULATE2
VAR_IN_OUT
	AXIS : Axis_REf;
END_VAR
END_METHOD

METHOD FILTERSTARTCONDITION
VAR_INPUT
	LRSETPOS : LREAL;
	LRSETVEL : LREAL;
	LRSETACC : LREAL;
END_VAR
VAR_IN_OUT
	AXIS : Axis_ref;
END_VAR
END_METHOD

METHOD GETOFFSETVALUES
VAR_OUTPUT
	LROFFSETPOS : LREAL;
	LROFFSETVEL : LREAL;
	LROFFSETACC : LREAL;
END_VAR
END_METHOD

METHOD CALLFUNCTION
VAR_INPUT
	UIINPUTDATAIDX : UINT;
	UIOUTPUTDATAIDX : UINT;
END_VAR
END_METHOD

METHOD COPYINPUTS : BOOL
VAR_INPUT
	IDX : WORD;
END_VAR
END_METHOD

METHOD COPYOUTPUTS : BOOL
VAR_INPUT
	IDX : WORD;
END_VAR
END_METHOD

METHOD CHECKINPUTDATA2
VAR_IN_OUT
	AXIS : Axis_REf;
END_VAR
END_METHOD

(* ---- L_CT1P_ONLINEIDENTSTIFFMECHANICS.fb ---- *)
FUNCTION_BLOCK L_CT1P_ONLINEIDENTSTIFFMECHANICS EXTENDS L_CT1P_OnlineIdentStiffMechanics_internal
VAR_INPUT
	XENABLE : BOOL := FALSE;
	XRESTART : BOOL := TRUE;
	ESTARTMODE : L_CT1P_StartMode := L_CT1P_StartMode.AutoInit;
	LRSTARTINERTIA : LREAL := 0.001;
	LRSTARTVISCOUSFRICTION : LREAL := 0.001;
	LRSTARTCOULOMBFRICTION : LREAL := 0.001;
	LRSTARTCONSTANTTORQUE : LREAL := 0.0;
	LRTHRESHOLDVALUE : LREAL := 30.0;
END_VAR
VAR_OUTPUT
	XBUSY : BOOL;
	XERROR : BOOL;
	EERRORID : L_IE1P_Error;
	XVALIDALL : BOOL;
	XVALIDINERTIA : BOOL;
	XVALIDVISCOUSFRICTION : BOOL;
	XVALIDCOULOMBFRICTION : BOOL;
	XVALIDCONSTANTTORQUE : BOOL;
	LRIDENTVELOCITY : LREAL;
	LRIDENTINERTIA : LREAL;
	LRIDENTVISCOUSFRICTION : LREAL;
	LRIDENTCOULOMBFRICTION : LREAL;
	LRIDENTCONSTANTTORQUE : LREAL;
	LRCONVERGENCE : LREAL;
END_VAR
VAR_IN_OUT
	AXIS : AXIS_REF;
END_VAR
VAR
	FBBASE : L_MC1P_Template;
	LICHANDLING : L_IMHP_LLMHandling;
	LREXTVELOCITY_ : LREAL;
	XEXTVELOCITYUSED : BOOL;
	XEXTVELOCITYSET : BOOL;
	EIDENTMODE : L_CT1P_IdentMode := L_CT1P_IdentMode.IdentAll;
	_MCCALL : L_UM1P_MCCall;
	_INPUTDATA : ARRAY [1..2] OF L_CT1P_OnlineIdentStiffMechanicsDoubleInput;
	_OUTPUTDATA : ARRAY [1..2] OF L_CT1P_OnlineIdentStiffMechanicsDoubleOutput;
	LREXTVELOCITY : LREAL;
END_VAR
END_FUNCTION_BLOCK

METHOD CALLFUNCTION
VAR_INPUT
	UIINPUTDATAIDX : UINT;
	UIOUTPUTDATAIDX : UINT;
END_VAR
END_METHOD

METHOD COPYINPUTS : BOOL
VAR_INPUT
	IDX : WORD;
END_VAR
END_METHOD

METHOD COPYOUTPUTS : BOOL
VAR_INPUT
	IDX : WORD;
END_VAR
END_METHOD

METHOD FUNCTIONWASCALLEDTWICE : BOOL
VAR_INPUT
	IDX : WORD;
END_VAR
END_METHOD

METHOD HANDLESTANDARDCALL : BOOL
END_METHOD

METHOD SYNCOUTPUTS
VAR_INPUT
	UICOPYOUTPUTFROMIDX : UINT;
	UICOPYOUTPUTTOIDX : UINT;
END_VAR
END_METHOD

METHOD COPYINPUTSINTERNAL
VAR_INPUT
	IDX : WORD;
END_VAR
END_METHOD

METHOD COPYOUTPUTSINTERNAL
VAR_INPUT
	IDX : WORD;
END_VAR
END_METHOD

METHOD RESETOUTPUTS
VAR_INPUT
	IDX : WORD;
END_VAR
END_METHOD

(* ---- L_CT1P_ONLINEIDENTSTIFFMECHANICS_INTERNAL.fb ---- *)
FUNCTION_BLOCK L_CT1P_ONLINEIDENTSTIFFMECHANICS_INTERNAL
VAR
	XREINIT_INT : BOOL := TRUE;
	EINITPARAMSOURCE_INT : L_CT1P_StartMode := L_CT1P_StartMode.AutoInit;
	LRINERTIAINIT_INT : LREAL := 0.001;
	LRCOULOMBFRICTIONINIT_INT : LREAL := 0.001;
	LRVISCOUSFRICTIONINIT_INT : LREAL := 0.001;
	LRCONSTANTTORQUEINIT_INT : LREAL := 0.0;
	EIDENTMODE_INT : L_CT1P_IdentMode := L_CT1P_IdentMode.IdentAll;
	LRTHRESHOLDVALUE_INT : LREAL := 30.0;
	LRVELOCITYIDENT_INT : LREAL;
	LRINERTIAIDENTKGCM2_INT : LREAL;
	LRVISCOUSDAMPINGIDENT_INT : LREAL;
	LRCONSTANTTORQUEIDENT_INT : LREAL;
	LRIDENTCOULOMBFRICTION_INT : LREAL;
	LRCONVERGENCE_INT : LREAL;
	XVALIDALL_INT : BOOL;
	XVALIDINERTIA_INT : BOOL;
	XVALIDVISCOUSDAMPING_INT : BOOL;
	XVALIDCONSTANTTORQUE_INT : BOOL;
	XVALIDCOULOMBFRICTION_INT : BOOL;
	XVALIDVISCOUSGRADIENT : BOOL;
	XVALIDCOULOMBGRADIENT : BOOL;
	XERROR_INT : BOOL;
	EERRORID_INT : L_IE1P_Error;
	PAXISREAL1 : POINTER TO _AXIS_REF_REAL;
	PAXISREAL2 : POINTER TO _AXIS_REF_REAL;
	XPARAMREADY : BOOL;
	XENABLEOLD : BOOL;
	XREINITOLD : BOOL;
	XREINITPULSE : BOOL;
	XREINITAFTERSTANDSTILL : BOOL;
	DICOUNTPLAUSIBILITYFAIL : DINT;
	DICOUNTPLAUSIBILITYFAILMAX : DINT;
	ICOUNTPLAUSIBILITYINITIALCHECK : INT;
	ILIMITNOPLAUSIBILITYREACHED_ : INT := 20000;
	LRTIMEPLAUSIBILITYFAILMAX_ : LREAL := 3.0;
	ICOUNTPLAUSIBILITYSUCCESS : INT;
	ILIMITPLAUSIBILITYSUCCESS_ : INT := 2000;
	XPLAUSIBILITYREACHED : BOOL;
	XDETECTPLAUSIBILITYFAIL : BOOL;
	LRTIMESTANDSTILLMAX_ : LREAL := 0.0;
	LRTIMECONSTANTVELOCITYMAX_ : LREAL := 5.0;
	LRVELSTANDSTILL_ : LREAL := 20.0;
	XSETVELSTANDSTILL : BOOL := FALSE;
	ICASEEXCITATION : INT;
	ICOUNTACCELERATION : INT := -1;
	INUMCOUNTSEXCIATIONMAX_ : INT := 10000;
	INUMCOUNTSEXCIATIONMIN_ : INT := 2000;
	LREXCITATIONPERCENTLIMIT_ : LREAL := 0.5;
	LRNOEXCITATIONPERCENTAGE : LREAL;
	LRTIMEMINLACKEXCITATION_ : LREAL := 1.0;
	AIEXCITATIONTIMES : ARRAY [0..1, 0..(ciLength - 1)] OF INT;
	IEXCITATIONBUFFERACT : INT;
	IEXCITATIONBUFFERSTART : INT;
	IEXCITATIONCOUNTALL : INT;
	IEXCITATIONCOUNT : INT;
	ICOUNTNOEXCITATION : INT;
	XDETECTLACKEXCITATION : BOOL;
	XWARNINGEXCITATIONFUNC : BOOL;
	ICOUNTSTANDSTILL : INT := -1;
	ICOUNTSTANDSTILLMAX : INT;
	ICOUNTCONSTANTVELOCITY : INT := -1;
	ICOUNTCONSTANTVELOCITYMAX : INT;
	XDETECTSTANDSTILL : BOOL;
	XDETECTSTANDSTILL_OLD : BOOL;
	XDETECTCONSTANTVELOCITY : BOOL;
	XDETECTCONSTANTVELOCITY_OLD : BOOL;
	LRJ_MOTOR1 : LREAL;
	LRJ_MOTOR2 : LREAL;
	LRNNENNMOTOR1 : LREAL := 3000.0;
	LRNNENNMOTOR2 : LREAL := 3000.0;
	LRRATIO1 : LREAL := 1;
	LRRATIO2 : LREAL := 1;
	LREXTVELOCITY1_LOCAL : LREAL;
	LREXTVELOCITY2_LOCAL : LREAL;
	LRINERTIAINITINTERN1 : LREAL := 0.001;
	LRINERTIAINITINTERN2 : LREAL := 0.001;
	LRVISCOUSDAMPINGINITINTERN1 : LREAL := 0.001;
	LRVISCOUSDAMPINGINITINTERN2 : LREAL := 0.001;
	LRCOULOMBDAMPINGINITINTERN1 : LREAL := 0.001;
	LRCOULOMBDAMPINGINITINTERN2 : LREAL := 0.001;
	LRCONSTANTTORQUEINITINTERN1 : LREAL := 0.0;
	LRCONSTANTTORQUEINITINTERN2 : LREAL := 0.0;
	LRINERTIAINITFACT1 : LREAL := 20;
	LRINERTIAINITFACT2 : LREAL := 5;
	LRINERTIAINITFACTFBINPUTS1 : LREAL := 1.5;
	LRINERTIAINITFACTFBINPUTS2 : LREAL := 0.5;
	LRFILTERTIME_XVALID : LREAL := 5000;
	LRFILTERCOUNTMAX : LREAL;
	LRINVFILTERCOUNTMAX : LREAL;
	LRVISCOUSGRADIENTVALIDCNT : LREAL;
	LRCOULOMBGRADIENTVALIDCNT : LREAL;
	LRGRADIENTCYCLECOUNT : LREAL;
	LRGRADIENTVALIDCOUNTMAX : LREAL;
	LRGRADIENTCYCLECOUNTMAX_ : LREAL := 10;
	LRGRADIENTTOLERANCE_ : LREAL := 5.0;
	LRGRADIENTVALIDTIME_ : LREAL := 5000;
	LRINERTIAIDENT_MEAN : LREAL;
	LRVISDAMPINGIDENT_MEAN : LREAL;
	LRCONSTORQUEIDENT_MEAN : LREAL;
	LRIDENTCOULOMBFRICTION_MEAN : LREAL;
	LRINERTIAIDENT_DIFF : LREAL;
	LRVISDAMPINGIDENT_DIFF : LREAL;
	LRCONSTORQUEIDENT_DIFF : LREAL;
	LRIDENTCOULOMBFRICTION_DIFF : LREAL;
	SCFRICTIONHIST : L_CT1P_FrictionHist;
	LRPT1FILTERTIMEINERTIA : LREAL := 5000;
	LRPT1FILTERTIMENORMINERTIA : LREAL;
	LRPT1FILTERTIMEDAMPING : LREAL := 5000;
	LRPT1FILTERTIMENORMDAMPING : LREAL;
	LRPT1FILTERTIMECONSTTORQUE : LREAL := 100;
	LRPT1FILTERTIMENORMCONSTTORQUE : LREAL;
	LRPT1FILTERTIMECOULOMBFRICTION : LREAL := 5000;
	LRPT1FILTERTIMENORMCOULOMBFRICTION : LREAL;
	LRPT1FILTERCONVERGENCE : LREAL := 1000;
	LRPT1FILTERNORMCONVERGENCE : LREAL;
	LRINERTIAVALIDCNT : LREAL;
	LRVISDAMPINGVALIDCNT : LREAL;
	LRCONSTORQUEVALIDCNT : LREAL;
	LRCOULOMBFRICTIONVALIDCNT : LREAL;
	LRVORSCHUBK1 : LREAL := 1;
	LRVORSCHUBK2 : LREAL := 1;
	LRM_IST_NORM : LREAL;
	LROMEGA_IST_NORM : LREAL;
	LRREFTORQUESCALING : LREAL;
	LRRATEDSPEEDSCALING : LREAL;
	LRINVREFTORQUESCALING : LREAL;
	LRINVRATEDSPEEDSCALING : LREAL;
	KALMANFILTER1 : L_CT1P_KalmanFilter_internal;
	KALMANFILTER2 : L_CT1P_KalmanFilter_internal;
	LRTORQUEINT1 : LREAL;
	LRTORQUEINT2 : LREAL;
	CILENGTH : INT := 30;
	LRGRADIENTCYCLECOUNTMAX : LREAL;
	LRGRADIENTTOLERANCE : LREAL;
	LRGRADIENTVALIDTIME : LREAL;
	LRTIMECONSTANTVELOCITYMAX : LREAL;
	LRTIMESTANDSTILLMAX : LREAL;
	LRTIMEVALIDFLAGS : LREAL;
	LRVELSTANDSTILL : LREAL;
END_VAR
END_FUNCTION_BLOCK

METHOD CALCSCALINGVALUES : BOOL
END_METHOD

METHOD CHECKPLAUSIBILITY : BOOL
END_METHOD

METHOD DETECTCONSTANTVELOCITY : BOOL
END_METHOD

METHOD DETECTLACKEXCITATION : BOOL
END_METHOD

METHOD DETECTPLAUSIBILITYFAIL
END_METHOD

METHOD DETECTSTANDSTILL : BOOL
END_METHOD

METHOD EVALUATEFRICTIONGRADIENT : BOOL
VAR_OUTPUT
	XVALIDVISCOUSGRADIENT : BOOL;
	XVALIDCOULOMBGRADIENT : BOOL;
END_VAR
END_METHOD

METHOD GENERATEOUTPUTSIGNALS
VAR_INPUT
	XSETOUTPDIRECT : BOOL;
END_VAR
END_METHOD

METHOD ONLINEIDENTSTIFFMECHANICS_INTERNAL
END_METHOD

METHOD READPARAM : BOOL
VAR_INPUT
	PAXISREAL : POINTER TO _AXIS_REF_REAL;
END_VAR
VAR_OUTPUT
	LRJ_MOTOR : LREAL;
	LRNNENNMOTOR : LREAL;
	LRVORSCHUBK : LREAL;
	LRRATIO : LREAL;
END_VAR
END_METHOD

METHOD SETIDENTMODE : BOOL
VAR_INPUT
	EIDENTMODE_INT : L_CT1P_IdentMode;
END_VAR
END_METHOD

METHOD SETQMATRIX : BOOL
VAR_INPUT
	LRQ_VALUE_00 : LREAL;
	LRQ_VALUE_06 : LREAL;
	LRQ_VALUE_12 : LREAL;
	LRQ_VALUE_18 : LREAL;
	LRQ_VALUE_24 : LREAL;
END_VAR
END_METHOD

METHOD COUNTLACKEXCITATION
VAR_INPUT
	ICURRENTCOUNT : INT;
END_VAR
END_METHOD

METHOD RESETEXCITATION
END_METHOD

METHOD UPDATESTARTACTBUFFER
END_METHOD

(* ---- L_CT1P_ONLINEIDENTSTIFFMECHANICSDOUBLE.fb ---- *)
FUNCTION_BLOCK L_CT1P_ONLINEIDENTSTIFFMECHANICSDOUBLE EXTENDS L_CT1P_OnlineIdentStiffMechanics_internal
VAR_INPUT
	XENABLE : BOOL := FALSE;
	XRESTART : BOOL := TRUE;
	ESTARTMODE : L_CT1P_StartMode := L_CT1P_StartMode.AutoInit;
	LRSTARTINERTIA : LREAL := 0.001;
	LRSTARTVISCOUSFRICTION : LREAL := 0.001;
	LRSTARTCOULOMBFRICTION : LREAL := 0.001;
	LRSTARTCONSTANTTORQUE : LREAL := 0.0;
	LRTHRESHOLDVALUE : LREAL := 30.0;
END_VAR
VAR_OUTPUT
	XBUSY : BOOL;
	XERROR : BOOL;
	EERRORID : L_IE1P_Error;
	XVALIDALL : BOOL;
	XVALIDINERTIA : BOOL;
	XVALIDVISCOUSFRICTION : BOOL;
	XVALIDCOULOMBFRICTION : BOOL;
	XVALIDCONSTANTTORQUE : BOOL;
	LRIDENTVELOCITY : LREAL;
	LRIDENTINERTIA : LREAL;
	LRIDENTVISCOUSFRICTION : LREAL;
	LRIDENTCOULOMBFRICTION : LREAL;
	LRIDENTCONSTANTTORQUE : LREAL;
	LRCONVERGENCE : LREAL;
END_VAR
VAR_IN_OUT
	AXIS1 : AXIS_REF;
	AXIS2 : AXIS_REF;
END_VAR
VAR
	FBBASE1 : L_MC1P_Template;
	FBBASE2 : L_MC1P_Template;
	LICHANDLING : L_IMHP_LLMHandling;
	LREXTVELOCITY1_ : LREAL;
	LREXTVELOCITY2_ : LREAL;
	XEXTVELOCITYUSED1 : BOOL;
	XEXTVELOCITYSET1 : BOOL;
	XEXTVELOCITYUSED2 : BOOL;
	XEXTVELOCITYSET2 : BOOL;
	EIDENTMODE : L_CT1P_IdentMode := L_CT1P_IdentMode.IdentAll;
	_MCCALL : L_UM1P_MCCall;
	_INPUTDATA : ARRAY [1..2] OF L_CT1P_OnlineIdentStiffMechanicsDoubleInput;
	_OUTPUTDATA : ARRAY [1..2] OF L_CT1P_OnlineIdentStiffMechanicsDoubleOutput;
	LREXTVELOCITY1 : LREAL;
	LREXTVELOCITY2 : LREAL;
END_VAR
END_FUNCTION_BLOCK

METHOD CALLFUNCTION
VAR_INPUT
	UIINPUTDATAIDX : UINT;
	UIOUTPUTDATAIDX : UINT;
END_VAR
END_METHOD

METHOD COPYINPUTS : BOOL
VAR_INPUT
	IDX : WORD;
END_VAR
END_METHOD

METHOD COPYOUTPUTS : BOOL
VAR_INPUT
	IDX : WORD;
END_VAR
END_METHOD

METHOD FUNCTIONWASCALLEDTWICE : BOOL
VAR_INPUT
	IDX : WORD;
END_VAR
END_METHOD

METHOD HANDLESTANDARDCALL : BOOL
END_METHOD

METHOD SYNCOUTPUTS
VAR_INPUT
	UICOPYOUTPUTFROMIDX : UINT;
	UICOPYOUTPUTTOIDX : UINT;
END_VAR
END_METHOD

METHOD COPYINPUTSINTERNAL
VAR_INPUT
	IDX : WORD;
END_VAR
END_METHOD

METHOD COPYOUTPUTSINTERNAL
VAR_INPUT
	IDX : WORD;
END_VAR
END_METHOD

(* ---- L_CT1P_OSCILLATIONCOMP.fb ---- *)
FUNCTION_BLOCK L_CT1P_OSCILLATIONCOMP EXTENDS L_MC1P_SetSetValueManipulator
VAR_INPUT
	XCONTINIOUSUPDATE : BOOL;
	LRAMPRATIO : LREAL := 1;
	LREIGENFREQ : LREAL := 0;
	ECOMPMODE : L_CT1P_OscCompMode;
	XMANIPULATETORQUE : BOOL;
END_VAR
VAR_OUTPUT
	XINEQOUT : BOOL;
END_VAR
VAR
	LICHANDLING : L_IMHP_LLMHandling;
	LRFDSET : LREAL;
	LRFDACT : LREAL;
	LRDFDACT : LREAL;
	LRDDFDACT : LREAL;
	LRDSET : LREAL;
	LRDACT : LREAL;
	LRDDACT : LREAL;
	LRDDDACT : LREAL;
	ECOMPMODEINT : L_CT1P_OscCompModeAct;
	LRCOEFFBLENDFACTORSET : LREAL;
	LRCOEFFBLENDFACTORACT : LREAL;
	LRDCOEFFBLENDFACTORACT : LREAL;
	LRDDCOEFFBLENDFACTORACT : LREAL;
	XCONTINIOUSUPDATEINT : BOOL;
	XMANIPULATETORQUEINT : BOOL;
	LRHOMINGOFFSETACT : LREAL;
	ALRFILTERCOEFF : ARRAY [1..3] OF LREAL;
	ALRDFILTERCOEFF : ARRAY [1..3] OF LREAL;
	ALRDDFILTERCOEFF : ARRAY [1..3] OF LREAL;
	ALRPOSBUFFER : ARRAY [1..cwBufferSize] OF LREAL;
	ALRVELBUFFER : ARRAY [1..cwBufferSize] OF LREAL;
	ALRACCBUFFER : ARRAY [1..cwBufferSize] OF LREAL;
	ALRTORQUEBUFFER : ARRAY [1..cwBufferSize] OF LREAL;
	ADIBUFFERINDEX : ARRAY [1..5] OF DINT;
	LRWEIGHTEDPOS : LREAL;
	LRWEIGHTEDVEL : LREAL;
	LRWEIGHTEDACC : LREAL;
	LRWEIGHTEDTORQUE : LREAL;
	DI1HALFPERIOD : DINT;
	DI2HALFPERIOD : DINT;
	LRHALFPERIOD : LREAL;
	LRSUBCYCLE1HALFPERIOD : LREAL;
	LRSUBCYCLE2HALFPERIOD : LREAL;
	UIINEQOUTCNT : UINT;
	DWACTFILTERDEPTH : DWORD;
	LRSETPOSINOLD : LREAL;
	LRSETVELINOLD : LREAL;
	LRSETACCINOLD : LREAL;
	LRSETTORQUEINOLD : LREAL;
	LRPOSOUTOLD : LREAL;
	LRVELOUTOLD : LREAL;
	LRACCOUTOLD : LREAL;
	LRTORQUEOUTOLD : LREAL;
	LRNUMMEMSIZEOLD : LREAL;
	XINEQOUTOLD : BOOL;
	LRMAXCHANGELRFD : LREAL := 0.0003;
	LRMAXCHANGELRD : LREAL := 0.0005;
	LRMAXCHANGEBLENDCOEFFS : LREAL := 0.0005;
	UIFILTERTIMELRFD : UINT := 10;
	UIFILTERTIMELRD : UINT := 10;
	UIMINLIMITERCYCLESFD : UINT := 50;
	UIMINLIMITERCYCLESD : UINT := 50;
	RATELIMITERFD : L_CT1P_RateLimiterCubicAvrgFilt;
	RATELIMITERD : L_CT1P_RateLimiterCubicAvrgFilt;
	RATELIMITERCOEFF : L_CT1P_RateLimiterCubicQuintic;
	XERROR_CHECKINPUTDATA : BOOL;
	DWSTANDSTILLCNT : DWORD;
	FBOCBASE : L_CT1P_OscillationCompBase;
	CWBUFFERSIZE : WORD := 2528;
	LRFDMIN : LREAL := 0.4;
	LRFDMAX : LREAL := 40;
	_CUSTOMINPUTDATA : ARRAY [1..2] OF L_CT1P_OscillationCompInput;
	_CUSTOMOUTPUTDATA : ARRAY [1..2] OF L_CT1P_OscillationCompOutput;
	_PCUSTOMINPUTDATA : POINTER TO L_CT1P_OscillationCompInput;
	_PCUSTOMOUTPUTDATA : POINTER TO L_CT1P_OscillationCompOutput;
	RATELIMPARA_COMPMODE : LREAL;
	RATELIMPARA_LRAMPRATIO : LREAL;
	RATELIMPARA_LREIGENFREQ : LREAL;
END_VAR
END_FUNCTION_BLOCK

METHOD CALLCYCLIC2
VAR_IN_OUT
	AXIS : AXIS_REF;
END_VAR
END_METHOD

METHOD READINPUTS2
VAR_IN_OUT
	AXIS : AXIS_REF;
END_VAR
END_METHOD

METHOD RESETOUTPUTS2
VAR_IN_OUT
	AXIS : Axis_REf;
END_VAR
END_METHOD

METHOD CALCULATE2
VAR_IN_OUT
	AXIS : Axis_REf;
END_VAR
END_METHOD

METHOD ENABLEEXIT2
VAR_IN_OUT
	AXIS : Axis_REf;
END_VAR
END_METHOD

METHOD ENABLEINIT2
VAR_IN_OUT
	AXIS : Axis_REf;
END_VAR
END_METHOD

METHOD LOADOFFSET2
VAR_INPUT
	OFFSET : LREAL;
END_VAR
VAR_IN_OUT
	AXIS : Axis_REf;
END_VAR
END_METHOD

METHOD RESET2
VAR_IN_OUT
	AXIS : Axis_REf;
END_VAR
END_METHOD

METHOD CALLFUNCTION
VAR_INPUT
	UIINPUTDATAIDX : UINT;
	UIOUTPUTDATAIDX : UINT;
END_VAR
END_METHOD

METHOD COPYINPUTS : BOOL
VAR_INPUT
	IDX : WORD;
END_VAR
END_METHOD

METHOD COPYOUTPUTS : BOOL
VAR_INPUT
	IDX : WORD;
END_VAR
END_METHOD

METHOD CALCFILTERVALUES
VAR_IN_OUT
	AXIS : AXIS_REF;
END_VAR
END_METHOD

METHOD CHECKINPUTDATA
END_METHOD

METHOD UPDATESYSTEMPARAMETER
VAR_IN_OUT
	AXIS : AXIS_REF;
END_VAR
END_METHOD

METHOD CALCWEIGTHEDDELTA
VAR_IN_OUT
	AXIS : Axis_REf;
END_VAR
END_METHOD

METHOD PRELOADARRAYS
END_METHOD

METHOD SHIFTINDICES
END_METHOD

(* ---- L_CT1P_OSCILLATIONCOMPBASE.fb ---- *)
FUNCTION_BLOCK L_CT1P_OSCILLATIONCOMPBASE
VAR
	LRREMVIB : LREAL := 0.1;
END_VAR
END_FUNCTION_BLOCK

METHOD CALCDAMPING : BOOL
VAR_INPUT
	LRAMPRATIO : LREAL;
END_VAR
VAR_OUTPUT
	LRDSET : LREAL;
END_VAR
END_METHOD

METHOD CALCFILTERVALUESBASE
VAR_INPUT
	ECOMPMODEINT : L_CT1P_OscCompModeAct;
	ALRFILTERCOEFF : REFERENCE TO ARRAY [1..3] OF LREAL;
	ALRDFILTERCOEFF : REFERENCE TO ARRAY [1..3] OF LREAL;
	ALRDDFILTERCOEFF : REFERENCE TO ARRAY [1..3] OF LREAL;
	LRDACT : LREAL;
	LRDDACT : LREAL;
	LRDDDACT : LREAL;
END_VAR
END_METHOD

METHOD CALCFILTERVALUES_ZV
VAR_INPUT
	LRDACT : LREAL;
	LRDDACT : LREAL;
	LRDDDACT : LREAL;
END_VAR
VAR_IN_OUT
	ZV : ARRAY [1..2, 1..3] OF LREAL;
END_VAR
END_METHOD

METHOD CALCFILTERVALUES_ZVD
VAR_INPUT
	LRDACT : LREAL;
	LRDDACT : LREAL;
	LRDDDACT : LREAL;
END_VAR
VAR_IN_OUT
	ZVD : ARRAY [1..3, 1..3] OF LREAL;
END_VAR
END_METHOD

(* ---- L_CT1P_PARAUTOTUNING.fb ---- *)
FUNCTION_BLOCK L_CT1P_PARAUTOTUNING EXTENDS L_CT1P_ParAutoTuninginternal
VAR_INPUT
	XENABLE : BOOL;
	AUTOTUNING : REFERENCE TO L_CT1P_Autotuning;
END_VAR
END_FUNCTION_BLOCK

(* ---- L_CT1P_PARAUTOTUNINGINTERNAL.fb ---- *)
FUNCTION_BLOCK L_CT1P_PARAUTOTUNINGINTERNAL
VAR_INPUT
	LRMAXVELOCITYDURINGSTANDSTILLRATIO_PCT : LREAL := 10.0;
	LRPROFILEVELOCITYRATIO_PCT : LREAL := 10.0;
	LRVPNINITFACTORMOTORINERTIA_PCT : LREAL := 100.0;
	LRVPNINITFACTORLOADINERTIA_PCT : LREAL := 25.0;
	LRVPNSTEPFACTOR_PCT : LREAL := 100.0;
	LRTNNINITFACTOR_PCT : LREAL := 100.0;
	LRVPPINITFACTOR_PCT : LREAL := 20.0;
	LRVPPSTEPFACTOR_PCT : LREAL := 100.0;
	LRSTARTMOVEMENTINPOSITIONTIMEOUT : LREAL := 10.0;
	WAUTOTUNEVPNCRITERIA : WORD := 1;
	WAUTOTUNETNNCRITERIA : WORD := 1;
	WAUTOTUNEVPPCRITERIA : WORD := 2;
	XUSE_0X2DE0_019_FORVELOCITYERROR : BOOL := FALSE;
END_VAR
END_FUNCTION_BLOCK

(* ---- L_CT1P_PLANECOMP.fb ---- *)
FUNCTION_BLOCK L_CT1P_PLANECOMP EXTENDS L_MC1P_CompensationBase
VAR_INPUT
	ALRBASE1POSITION : POINTER TO LREAL;
	ALRBASE2POSITION : POINTER TO LREAL;
	ALRAXISCORRECTION : POINTER TO LREAL;
END_VAR
VAR_OUTPUT
	LRACTCORRECTION : LREAL;
END_VAR
VAR_IN_OUT
	BASE1 : AXIS_REF;
	BASE2 : AXIS_REF;
END_VAR
VAR
	LICHANDLING : L_IMHP_LLMHandling;
	LRCORRECTIONPOS : LREAL;
	LRCORRECTIONVEL : LREAL;
	LRCORRECTIONACC : LREAL;
	LRCORRECTIONPOSOLD : LREAL;
	LRCORRECTIONVELOLD : LREAL;
	UDINBROFXVALUES : UDINT;
	UDINBROFYVALUES : UDINT;
	XFIRSTCALL : BOOL;
	_CUSTOMINPUTDATA : ARRAY [1..2] OF L_CT1P_PlaneCompInput;
	_CUSTOMOUTPUTDATA : ARRAY [1..2] OF L_CT1P_PlaneCompOutput;
	_PCUSTOMINPUTDATA : POINTER TO L_CT1P_PlaneCompInput;
	_PCUSTOMOUTPUTDATA : POINTER TO L_CT1P_PlaneCompOutput;
	_ITFBASE1 : L_MC1P_IAXIS_REF_MASTERVALUES;
	_ITFBASE2 : L_MC1P_IAXIS_REF_MASTERVALUES;
END_VAR
END_FUNCTION_BLOCK

METHOD CALLCYCLIC2
VAR_IN_OUT
	AXIS : Axis_REf;
END_VAR
END_METHOD

METHOD CHECKINPUTDATA2
VAR_IN_OUT
	AXIS : Axis_REf;
END_VAR
END_METHOD

METHOD READINPUTS2
VAR_IN_OUT
	AXIS : Axis_REf;
END_VAR
END_METHOD

METHOD RESETOUTPUTS2
VAR_IN_OUT
	AXIS : Axis_REf;
END_VAR
END_METHOD

METHOD CALCULATE2
VAR_IN_OUT
	AXIS : Axis_REf;
END_VAR
END_METHOD

METHOD FILTERSTARTCONDITION
VAR_INPUT
	LRSETPOS : LREAL;
	LRSETVEL : LREAL;
	LRSETACC : LREAL;
END_VAR
VAR_IN_OUT
	AXIS : Axis_ref;
END_VAR
END_METHOD

METHOD GETOFFSETVALUES
VAR_OUTPUT
	LROFFSETPOS : LREAL;
	LROFFSETVEL : LREAL;
	LROFFSETACC : LREAL;
END_VAR
END_METHOD

METHOD CALLFUNCTION
VAR_INPUT
	UIINPUTDATAIDX : UINT;
	UIOUTPUTDATAIDX : UINT;
END_VAR
END_METHOD

METHOD COPYINPUTS : BOOL
VAR_INPUT
	IDX : WORD;
END_VAR
END_METHOD

METHOD COPYOUTPUTS : BOOL
VAR_INPUT
	IDX : WORD;
END_VAR
END_METHOD

METHOD INDEX : UDINT
VAR_INPUT
	I : UDINT;
	J : UDINT;
	STRIDE : UDINT;
END_VAR
END_METHOD

METHOD PRV2DINTERPOLATION : BOOL
VAR_INPUT
	LRX : LREAL;
	LRY : LREAL;
END_VAR
VAR_OUTPUT
	XERROR : BOOL;
	EERRORID : L_IE1P_Error;
	LRZ : LREAL;
END_VAR
END_METHOD

(* ---- L_CT1P_PROCESSCONTROLLER.fb ---- *)
FUNCTION_BLOCK L_CT1P_PROCESSCONTROLLER
VAR_INPUT
	LRSETVALUE : LREAL := 0.0;
	XLOADACTVALUE : BOOL := FALSE;
	LRACTVALUE : LREAL := 0.0;
	LRDELAYTIME : LREAL := 0.001;
	LRGAIN : LREAL := 1.0;
	LRGAINADAPT : LREAL := 0.0;
	LRRESETTIME : LREAL := 1.0;
	LRRATETIME : LREAL := 0.0;
	XRESET : BOOL := FALSE;
	XLOADINTVALUE : BOOL := FALSE;
	LRINTVALUE : LREAL := 0.0;
	LRACC : LREAL := 0.0;
	LRDEC : LREAL := 0.0;
	LRINFLUENCE : LREAL := 0.0;
	LRREDRANGE : LREAL := 0.0;
	LRREDGAIN : LREAL := 0.0;
	LRPOSLIMITVALUE : LREAL := L_UMTP_Math.gC_POSITIVE_LIMIT_32BIT;
	LRNEGLIMITVALUE : LREAL := L_UMTP_Math.gC_NEGATIVE_LIMIT_32BIT;
	ALRXVALUES : ARRAY [1..5] OF LREAL := [5(0)];
	ALRYVALUES : ARRAY [1..5] OF LREAL := [1, 4(0)];
END_VAR
VAR_OUTPUT
	LROUT : LREAL;
	LROUTRED : LREAL;
	LRSETRAMPVALUEOUT : LREAL;
	LRDEVIATION : LREAL;
	XLIMITACTIVE : BOOL;
	XERROR : BOOL;
	EERRORID : L_IE1P_Error;
END_VAR
VAR
	LRTASKCYCLE : LREAL := -1.0;
	LRINVTASKCYCLE : LREAL;
	LRTIME : LREAL;
	LRACTDELAY : LREAL;
	LRDIFF : LREAL;
	LRDIFFOLD : LREAL;
	LRABSDIFF : LREAL;
	LRPTEMP : LREAL;
	LRITEMP : LREAL;
	LRDTEMP : LREAL;
	LRTEMP : LREAL;
	LRRESGAIN : LREAL;
	CURVE : L_USPP_Curve;
	RAMP : L_MC1P_HlpRampGenerator;
	LRINT : LREAL;
	IDX : WORD;
	XLOADPVALUE : BOOL;
	XLOADIVALUE : BOOL;
	XLOADDVALUE : BOOL;
	LRPVALUE : LREAL;
	LRIVALUE : LREAL;
	LRDVALUE : LREAL;
	WPIDMODE : WORD;
	PIDMODE : WORD;
END_VAR
END_FUNCTION_BLOCK

METHOD GAINFRAC
VAR_INPUT
	LRGAIN_N : LREAL;
	LRINT : LREAL;
	LRREM : LREAL;
END_VAR
END_METHOD

METHOD GET_DPROCESSCONTROLLEROUT : LREAL
END_METHOD

METHOD GET_IPROCESSCONTROLLEROUT : LREAL
END_METHOD

METHOD GET_PPROCESSCONTROLLEROUT : LREAL
END_METHOD

METHOD SET_DPROCESSCONTROLLEROUT
VAR_INPUT
	LRVALUE : LREAL;
END_VAR
END_METHOD

METHOD SET_IPROCESSCONTROLLEROUT
VAR_INPUT
	LRVALUE : LREAL;
END_VAR
END_METHOD

METHOD SET_PPROCESSCONTROLLEROUT
VAR_INPUT
	LRVALUE : LREAL;
END_VAR
END_METHOD

(* ---- L_CT1P_RATELIMITERCUBIC.fb ---- *)
FUNCTION_BLOCK L_CT1P_RATELIMITERCUBIC
VAR_INPUT
	XENABLE : BOOL;
	XPRELOADVALUE : BOOL;
	LRIN : LREAL;
	LRMAXCHANGEPERCYCLE : LREAL;
	UIMINLIMITERCYCLES : UINT := 10;
END_VAR
VAR_OUTPUT
	LROUT : LREAL;
	LRDOUT : LREAL;
	LRDDOUT : LREAL;
END_VAR
VAR
	LRIN_OLD : LREAL;
	ALRCOEFFS : ARRAY [0..3] OF LREAL;
	ALRCOEFFSINT : ARRAY [0..3] OF LREAL;
	XNEWCOEFFSVALID : BOOL;
	LRTBLENDINT : LREAL;
	LRTBLEND : LREAL;
	LRINVTBLEND : LREAL;
	LRBLENDIPOCOUNTER : LREAL;
	LRTMP1 : LREAL;
	LRTMP2 : LREAL;
	LRTMP3 : LREAL;
	LRTEXTREMA : LREAL;
	LROUTEXTREMA : LREAL;
	LRSIGN : LREAL;
END_VAR
END_FUNCTION_BLOCK

(* ---- L_CT1P_RATELIMITERCUBICAVRGFILT.fb ---- *)
FUNCTION_BLOCK L_CT1P_RATELIMITERCUBICAVRGFILT EXTENDS L_UBUP_MemoryProvider
VAR_INPUT
	XENABLE : BOOL;
	XPRELOADVALUE : BOOL;
	LRIN : LREAL;
	LRMAXCHANGEPERCYCLE : LREAL;
	UIFILTERTIME : UINT;
	UIMINLIMITERCYCLES : UINT := 10;
END_VAR
VAR_OUTPUT
	XERROR : BOOL;
	EERRORID : L_IE1P_Error;
	LROUT : LREAL;
	LRDOUT : LREAL;
	LRDDOUT : LREAL;
END_VAR
VAR
	LRTASKCYCLE : LREAL := -1;
	XENABLE_R : R_Trig;
	AMEM : ARRAY [1..2] OF ARRAY [1..cuiFilterSizeMax] OF LREAL;
	FB_AVG : L_USPP_AverageFilterRecursive;
	PXDUMMY : POINTER TO BOOL;
	RAMPCUB : L_CT1P_RateLimiterCubic;
	LRINOLD : LREAL;
	LRDIN : LREAL;
	CUIFILTERSIZEMAX : UINT := 31;
	PTR : POINTER TO BYTE;
	SIZE : UDINT;
END_VAR
END_FUNCTION_BLOCK

(* ---- L_CT1P_RATELIMITERCUBICQUINTIC.fb ---- *)
FUNCTION_BLOCK L_CT1P_RATELIMITERCUBICQUINTIC
VAR_INPUT
	XENABLE : BOOL;
	XPRELOADVALUE : BOOL;
	LRIN : LREAL;
	LRMAXCHANGEPERCYCLE : LREAL;
	UIMINLIMITERCYCLES : UINT := 10;
END_VAR
VAR_OUTPUT
	LROUT : LREAL;
	LRDOUT : LREAL;
	LRDDOUT : LREAL;
END_VAR
VAR
	LRIN_OLD : LREAL;
	ALRCOEFFS : ARRAY [0..5] OF LREAL;
	ALRCOEFFSINT : ARRAY [0..5] OF LREAL;
	XNEWCOEFFSVALID : BOOL;
	LRTBLENDINT : LREAL;
	LRTBLEND : LREAL;
	LRINVTBLEND : LREAL;
	LRBLENDIPOCOUNTER : LREAL;
	LRTMP1 : LREAL;
	LRTMP2 : LREAL;
	LRTMP3 : LREAL;
	LRTEXTREMA : LREAL;
	LROUTEXTREMA : LREAL;
	LRSIGN : LREAL;
	XPOLY5 : BOOL := TRUE;
END_VAR
END_FUNCTION_BLOCK

(* ---- L_CT1P_RATELIMITERLINEAR.fb ---- *)
FUNCTION_BLOCK L_CT1P_RATELIMITERLINEAR
VAR_INPUT
	XENABLE : BOOL;
	XPRELOADVALUE : BOOL;
	LRIN : LREAL;
	LRMAXCHANGEPERCYCLE : LREAL;
END_VAR
VAR_OUTPUT
	LROUT : LREAL;
	LRDOUT : LREAL;
	LRDDOUT : LREAL;
END_VAR
END_FUNCTION_BLOCK

(* ---- L_CT1P_TORQUEPRECONTROL.fb ---- *)
FUNCTION_BLOCK L_CT1P_TORQUEPRECONTROL EXTENDS L_MC1P_Template
VAR_INPUT
	XENABLE : BOOL;
	EPRECONTROLMODE : L_MC1P_PreControlMode := L_MC1P_PreControlMode.ExclusiveOffsetTorque;
	LRINERTIA : LREAL;
	LRVISCOUSFRICTION : LREAL;
	LRCOULOMBFRICTION : LREAL;
	LRCONSTANTTORQUE : LREAL;
	LRTORQUEOVERRIDE : LREAL := 1.0;
	LRTORQUELIMITFACTOR : LREAL := 1.0;
	LRTORQUERATELIMIT : LREAL := 0.0;
END_VAR
VAR_OUTPUT
	XBUSY : BOOL;
	XERROR : BOOL;
	EERRORID : L_IE1P_Error;
	LRSETTORQUEOUT : LREAL;
END_VAR
VAR
	LICHANDLING : L_IMHP_LLMHandling;
	PAXISREAL : POINTER TO _AXIS_REF_REAL;
	XENABLEOLD : BOOL;
	LRTORQUE_J : LREAL;
	LRTORQUE_VISCFRICTION : LREAL;
	LRTORQUE_COULFRIC : LREAL;
	LRTORQUEPRECONTROL : LREAL;
	LRTORQUEPRECONTROLNEW : LREAL;
	LRTORQUEDELTACYCLE : LREAL;
	LRTORQUELIMIT : LREAL;
	LRTMP : LREAL;
	L_MC1P_SETTORQUEOFFSET0 : L_MC1P_SetTorqueOffset;
	XUSEFILTEREDVALUES : BOOL := TRUE;
	LRSETACCELERATION : LREAL;
	LRSETVELOCITY : LREAL;
	LRVELMINCOULOMBFRICTION : LREAL := L_MC1P_Constants.gc_eps_real;
	LROVERRIDECOULOMBFRICTION : LREAL := 1.0;
	_MCCALL : L_UM1P_MCCall;
	_INPUTDATA : ARRAY [1..2] OF L_CT1P_TorquePreControlInput;
	_OUTPUTDATA : ARRAY [1..2] OF L_CT1P_TorquePreControlOutput;
	_PINPUTDATA : POINTER TO L_CT1P_TorquePreControlInput;
	_POUTPUTDATA : POINTER TO L_CT1P_TorquePreControlOutput;
	OVERRIDECOULOMBFRICTION : LREAL;
	USEFILTEREDVALUES : BOOL;
	VELMINCOULOMBFRICTION : LREAL;
END_VAR
END_FUNCTION_BLOCK

METHOD CALLFUNCTION
VAR_INPUT
	UIINPUTDATAIDX : UINT;
	UIOUTPUTDATAIDX : UINT;
END_VAR
END_METHOD

METHOD COPYINPUTS : BOOL
VAR_INPUT
	IDX : WORD;
END_VAR
END_METHOD

METHOD COPYOUTPUTS : BOOL
VAR_INPUT
	IDX : WORD;
END_VAR
END_METHOD

METHOD FUNCTIONWASCALLEDTWICE : BOOL
VAR_INPUT
	IDX : WORD;
END_VAR
END_METHOD

METHOD HANDLESTANDARDCALL : BOOL
END_METHOD

METHOD SYNCOUTPUTS
VAR_INPUT
	UICOPYOUTPUTFROMIDX : UINT;
	UICOPYOUTPUTTOIDX : UINT;
END_VAR
END_METHOD
